(* IEC 61131-3 sources: daoli-st-library/DL_Device (part 25) *)

(* ---- FB_DL_IvBcdExport.st ---- *)
(*==============================================================================
 * 组件名称 (Component)  : FB_DL_IvBcdExport
 * 所属子库 (Sublibrary) : DL_Device
 * 当前版本 (Version)    : 1.0.0
 * 兼容性   (Platform)   : CODESYS 3.5+ / TwinCAT 3 / 汇川 InoProShop / 施耐德 Machine Expert
 *                         仅依赖 Standard.library（TON / R_TRIG），零厂商私有库
 * 功能描述 (Function)   : IV 测试仪 BCD 拨码设定导出。
 *                         把上位下发的十进制设定值（0..9999）拆成四位十进制数字，打包成 BCD 字，
 *                         经"导出脉冲 → 等回读 → 逐位比对"的握手闭环确认测试仪已正确接收；
 *                         回读不一致或超时即锁存故障，等人工复位后重导。
 *                         **面板互转语义（双向，写死）**：
 *                           正解：value → 四位数字 d1(个)…d4(千) → uBcd = d4·16#1000 + d3·16#0100 + d2·16#0010 + d1
 *                           反解：uBcd → value（用于回读通道是 BCD 字的机型，本件按整值比对不拆位）
 *                         两位以上的半字节合法性由"十进制拆分"结构性保证（每位恒 0..9），
 *                         故不存在"非 BCD 半字节"可导出；真正的越界风险在**设定值本身越域**，
 *                         故设 0..9999 域闸 + 越域拒导出（eRangeBad，信息级，不锁存）。
 *                         验收向量：
 *                           ① 设定 1234 → 数字 d1=4, d2=3, d3=2, d4=1；uBcd = 16#1234
 *                           ② 设定 0    → 数字全 0；uBcd = 16#0000（合法边界，不拒算）
 *                           ③ 设定 9999 → uBcd = 16#9999（上界，不溢出）
 *                           ④ 设定 10000 → 拒导出 + eRangeBad（域闸，信息级）
 *                           ⑤ 回读 = 16#1234 → bReadbackOk；回读 = 16#1235 → 锁存 eRbMismatch
 * 接口     (Interface)  : 入 iSetValue 设定值、bExport 导出沿、bReadbackValid 回读有效、
 *                         iReadbackBcd 回读 BCD 字、tReadbackTo 回读超时、bReset 复位沿；
 *                         出 uBcdPacked 打包 BCD 字、abDigits 四位数字（1..4 = 个/十/百/千）、
 *                         bExported 导出脉冲（单拍）、bReadbackOk 回读一致脉冲（单拍）、
 *                         bRbFailed 回读失败锁存、eState 相、eCause 成因、bError 故障标志。
 * 边界     (Boundary)   : ① **属主边界（写死）：本件只做"设定值编码 + 导出握手"，不驱动拨码
 *                         继电器/光电隔离板、不解析 IV 测量曲线**（属测试仪通讯件与曲线件）；
 *                         ② **域闸**：iSetValue 越 0..9999 → 拒导出（信息级 eRangeBad，不锁存、
 *                         不改已导出值）；③ **移位量常量化**：打包移位量取常量 0/4/8/12，
 *                         恒小于 WORD 位宽 16，跨平台无未定义行为（R48/R295）；
 *                         ④ **回读超时 TON**：tonRb 段 0 无条件调用，IN 串 (NOT _bFault)，
 *                         故障期不累计，复位同拍不会立即重锁（R252）；
 *                         ⑤ **锁存解除式**：bRbFailed 与 eFault 仅由 bReset 上升沿解除
 *                         （R228B 唯一迁出），bReset 为外部引脚、恒可达；
 *                         ⑥ **握手单拍脉冲三律**：导出脉冲与回读成功脉冲均在 CASE 内用内部位
 *                         置位、段尾统一映射出口，禁同相内置位后同相撤位（R129）；
 *                         ⑦ 零全局耦合、零物理地址。
 * 分工声明 (Scope)      : 本件只管"设定值 BCD 导出与回读校验"。不接管：花篮标签打印联动
 *                         （属 FB_DL_CassetteBcdLabel）、纯数值 BCD 转换原子件（属 FC_DL_WordToBcd 族）、
 *                         IV 量测流程（属测试顺控件）。
 * 来源标签 (Source Tag) : ROADMAP 空勾真缺口 P2（BCD 设定导出，自研 clean-room）
 * 码表     (Codes)      : 本件不占用任何全局数字码位（零码位范式 R297）；诊断由 BOOL + ENUM 出口承担。
 * 红线自检 (Redline)    : R1 ✓ 零 GVL/VAR_EXTERNAL ｜ R2 ✓ 零 %I/%Q/%M ｜ R3 ✓ 纯 IEC 61131-3
 *                         R4 ✓ 域闸 + 常量移位 + 超时 TON + 单拍脉冲两段式 ｜ R5 ✓ 声明逐行同行双语注释
 *                         R6 ✓ ENUM+CASE 含 ELSE 兜底 ｜ R7 ✓ TON/R_TRIG 段 0 无条件刷新
 * 修订历史 (Revision)   : 2026-11-19  v1.0.0  R47 首版（批次 2 · 序号 10）
 *==============================================================================*)

TYPE E_DL_IbeState :
(
    eIdle    := 0,    // 待机相（可接受导出请求） / Idle, ready for an export request
    eWaitRead:= 10,   // 等回读相（握手窗口内） / Waiting for the read-back
    eFault   := 90    // 故障相（等复位） / Fault, awaiting reset
);
END_TYPE

TYPE E_DL_IbeCause :
(
    eNone       := 0,   // 无异常 / No anomaly
    eRangeBad   := 1,   // 设定值越 0..9999（信息级，拒导出） / Set point out of 0..9999, info level
    eRbMismatch := 2,   // 回读不一致（锁存，故障级） / Read-back mismatch, latched, fault level
    eRbTimeout  := 3,   // 回读超时（锁存，故障级） / Read-back timeout, latched, fault level
    eCfgIllegal := 4,   // 组态非法（超时非正） / Illegal configuration, non-positive timeout
    ePhaseBad   := 5    // 非法相位兜底 / Illegal phase fallback
);
END_TYPE

FUNCTION_BLOCK FB_DL_IvBcdExport
VAR_INPUT
    iSetValue     : INT := 0;              // 设定值，域 0..9999 [-] / Set point, domain 0..9999
    bExport       : BOOL := FALSE;         // 导出请求沿 [-] / Export request edge
    bReadbackValid: BOOL := FALSE;         // 回读有效（当拍电平） [-] / Read-back valid, level
    iReadbackBcd  : INT := 0;              // 回读 BCD 字（按整值比对） [BCD] / Read-back BCD word, compared as a whole
    tReadbackTo   : TIME := T#2S;          // 回读超时，域 > T#0S [ms] / Read-back timeout, > T#0S
    bReset        : BOOL := FALSE;         // 故障复位沿 [-] / Fault reset edge
END_VAR
VAR_OUTPUT
    uBcdPacked  : WORD := 16#0000;                       // 打包 BCD 字（千/百/十/个） [BCD] / Packed BCD word
    abDigits    : ARRAY[1..4] OF BYTE;                   // 四位十进制数字（1=个,2=十,3=百,4=千） [-] / Four decimal digits
    bExported   : BOOL := FALSE;                         // 导出脉冲（单拍） [-] / Export pulse, single scan
    bReadbackOk : BOOL := FALSE;                         // 回读一致脉冲（单拍） [-] / Read-back match pulse, single scan
    bRbFailed   : BOOL := FALSE;                         // 回读失败锁存（等复位） [-] / Read-back failure, latched
    eState      : E_DL_IbeState := E_DL_IbeState.eIdle;  // 相出口 [-] / Phase outlet
    eCause      : E_DL_IbeCause := E_DL_IbeCause.eNone;  // 成因出口（R190 归因唯一） [-] / Cause outlet
    bError      : BOOL := FALSE;                         // 故障标志（仅故障级成因） [-] / Error flag, fault level only
END_VAR
VAR
    _eState   : E_DL_IbeState := E_DL_IbeState.eIdle;    // 内部相（CASE 唯一写入目标） / Internal phase
    _eCause   : E_DL_IbeCause := E_DL_IbeCause.eNone;    // 成因锁存量 / Latched cause
    _bFault   : BOOL := FALSE;                           // 故障锁存位 / Latched fault bit
    _bRbFail  : BOOL := FALSE;                           // 回读失败锁存位 / Latched read-back failure
    _iWork    : INT := 0;                                // 十进制拆分工作值 [-] / Decimal split working value
    _uBcd     : WORD := 16#0000;                         // 打包工作值 [BCD] / Packing working value
    _iRbExp   : INT := 0;                                // 期望回读值（导出时的 BCD 整值） [BCD] / Expected read-back value
    _bExported: BOOL := FALSE;                           // 导出脉冲内部位（单拍） / Internal export pulse
    _bRbOk    : BOOL := FALSE;                           // 回读成功内部位（单拍） / Internal read-back OK pulse
    _bCfgBad  : BOOL := FALSE;                           // 组态非法当拍量 / Illegal configuration this scan
    tonRb     : TON;                                     // 回读超时实例，段 0 无条件调用 / Read-back timeout instance
    rtExport  : R_TRIG;                                  // 导出沿实例，段 0 无条件调用 / Export edge instance
    rtReset   : R_TRIG;                                  // 复位沿实例，段 0 无条件调用 / Reset edge instance
END_VAR
VAR CONSTANT
    DL_IBE_MAX  : INT := 9999;            // 设定值上限（四位十进制） [-] / Set-point upper bound
    DL_IBE_SH0  : WORD := 16#0000;        // 个位打包基准（占位常量，便于口径统一） [BCD] / Units packing base
    DL_IBE_SH4  : INT := 4;               // 十位左移量（恒 < 16，R48） [bit] / Tens shift, always below 16 bits
    DL_IBE_SH8  : INT := 8;               // 百位左移量（恒 < 16，R48） [bit] / Hundreds shift
    DL_IBE_SH12 : INT := 12;              // 千位左移量（恒 < 16，R48） [bit] / Thousands shift
    DL_IBE_MSK  : WORD := 16#000F;        // 半字节掩码（非事件码，头注释声明） [bit] / Nibble mask, not an event code
END_VAR

(* —— 段 0：组态闸 + TON 与两沿无条件周期刷新（R228A；IN 串故障否决，R252） —— *)
_bCfgBad := (tReadbackTo <= T#0S);                             // 回读超时须为正 / Timeout must be positive
rtExport(CLK := bExport);                                      // 导出沿 / Export edge
rtReset(CLK := bReset);                                        // 复位沿 / Reset edge
tonRb(IN := (_eState = E_DL_IbeState.eWaitRead) AND (NOT _bFault), PT := tReadbackTo);   // 回读超时（等回读相派生） / Read-back timeout

(* —— 段 1：单拍量预清零（锁存量 _eCause/_bFault/_bRbFail/_iRbExp 不入清单，R107） —— *)
_bExported := FALSE;                                           // 导出脉冲预清 / Export pulse preset
_bRbOk     := FALSE;                                           // 回读成功脉冲预清 / Read-back OK pulse preset
bError     := FALSE;                                           // 故障标志预清（R45 配对） / Error preset

(* —— 段 2：组态闸（非法即锁存故障级） —— *)
IF _bCfgBad THEN
    _eCause := E_DL_IbeCause.eCfgIllegal;                       // 归因：组态非法 / Cause: illegal configuration
    _bFault := TRUE;                                            // 锁存 / Latch
    _eState := E_DL_IbeState.eFault;                            // 入故障相 / Enter fault phase
END_IF

(* —— 段 3：迁出链（bReset 上升沿：清故障与回读失败锁存，R228B） —— *)
IF rtReset.Q THEN
    _bFault  := FALSE;                                          // 清故障锁存 / Clear fault latch
    _bRbFail := FALSE;                                          // 清回读失败锁存 / Clear read-back failure latch
    _eCause  := E_DL_IbeCause.eNone;                            // 清成因 / Clear cause
    _eState  := E_DL_IbeState.eIdle;                            // 回待机相 / Back to idle
END_IF

(* —— 段 4：相迁移（导出 / 回读握手闭环） —— *)
IF (NOT _bFault) AND (NOT _bCfgBad) THEN
    CASE _eState OF

    E_DL_IbeState.eIdle:
        IF rtExport.Q THEN
            IF (iSetValue < 0) OR (iSetValue > DL_IBE_MAX) THEN
                _eCause := E_DL_IbeCause.eRangeBad;              // 域闸：越域拒导出（信息级，不锁存） / Out of range, info level
            ELSE
                (* 十进制拆分（每位恒 0..9，半字节合法由构造保证） *)
                _iWork := iSetValue;                             // 取设定值 / Take the set point
                abDigits[1] := INT_TO_BYTE(_iWork MOD 10);       // 个位 / Units
                _iWork := _iWork / 10;                           // 去掉个位 / Drop the units digit
                abDigits[2] := INT_TO_BYTE(_iWork MOD 10);       // 十位 / Tens
                _iWork := _iWork / 10;                           // 去掉十位 / Drop the tens digit
                abDigits[3] := INT_TO_BYTE(_iWork MOD 10);       // 百位 / Hundreds
                _iWork := _iWork / 10;                           // 去掉百位 / Drop the hundreds digit
                abDigits[4] := INT_TO_BYTE(_iWork MOD 10);       // 千位 / Thousands

                (* 打包 BCD：移位量为常量，跨平台安全（R48/R295） *)
                _uBcd := SHL(BYTE_TO_WORD(abDigits[4]), DL_IBE_SH12)
                      OR SHL(BYTE_TO_WORD(abDigits[3]), DL_IBE_SH8)
                      OR SHL(BYTE_TO_WORD(abDigits[2]), DL_IBE_SH4)
                      OR (BYTE_TO_WORD(abDigits[1]) AND DL_IBE_MSK);
                uBcdPacked := _uBcd;                             // 打包字出口 / Packed word outlet
                _iRbExp := WORD_TO_INT(_uBcd);                   // 期望回读值（整值比对） / Expected read-back
                _bExported := TRUE;                              // 导出脉冲（内部位，段 7 映射） / Internal export pulse
                _eState := E_DL_IbeState.eWaitRead;              // 进等回读相 / Enter the wait-read phase
            END_IF
        END_IF

    E_DL_IbeState.eWaitRead:
        IF bReadbackValid THEN
            IF iReadbackBcd = _iRbExp THEN
                _bRbOk := TRUE;                                  // 回读一致（内部位） / Read-back matches
                _eState := E_DL_IbeState.eIdle;                  // 回待机相 / Back to idle
            ELSE
                _bRbFail := TRUE;                                // 回读不一致：锁存 / Mismatch: latch
                _bFault  := TRUE;                                // 故障锁存 / Latch the fault
                _eCause  := E_DL_IbeCause.eRbMismatch;           // 归因：回读不一致 / Cause: read-back mismatch
                _eState  := E_DL_IbeState.eFault;                // 入故障相 / Enter fault phase
            END_IF
        ELSIF tonRb.Q THEN
            _bRbFail := TRUE;                                    // 回读超时：锁存 / Timeout: latch
            _bFault  := TRUE;                                    // 故障锁存 / Latch the fault
            _eCause  := E_DL_IbeCause.eRbTimeout;                // 归因：回读超时 / Cause: read-back timeout
            _eState  := E_DL_IbeState.eFault;                    // 入故障相 / Enter fault phase
        END_IF

    E_DL_IbeState.eFault:
        ;                                                        // 故障相：仅等复位沿 / Wait for the reset edge only

    ELSE
        _eCause := E_DL_IbeCause.ePhaseBad;                      // 归因：非法相位 / Cause: illegal phase
        _bFault := TRUE;                                         // 锁存 / Latch
        _eState := E_DL_IbeState.eFault;                         // 强拉故障相 / Force fault phase

    END_CASE
END_IF

(* —— 段 5：出口单点映射（名实双出口，R191） —— *)
bExported   := _bExported;                                       // 导出脉冲出口 / Export pulse outlet
bReadbackOk := _bRbOk;                                           // 回读成功脉冲出口 / Read-back OK outlet
bRbFailed   := _bRbFail;                                         // 回读失败出口 / Read-back failure outlet
eState      := _eState;                                          // 相出口 / Phase outlet
eCause      := _eCause;                                          // 成因出口 / Cause outlet
bError      := _bFault;                                          // 故障标志 / Error flag

END_FUNCTION_BLOCK

(* ---- FB_DL_JunctionBoxPottingCheck.st ---- *)
(*
  FB_DL_JunctionBoxPottingCheck  —  接线盒灌胶量与固化判定 / Junction box potting quantity and cure check
  分类 Category : DL_Device
  码位 Code     : 16#03_2_14
  段位说明      : 03_2 段低半字节 00~0F 已满（05 为历史空穴留存），进位 14 段续号（R192）
  版本 Version  : 1.0.0
  来源 Source   : t2-1-lgf-technology — IEC 61131-3 标准语义的道莅防御性实现
  溯源 Origin   : clean-room 实现，灌胶积分与固化当量公开工艺语义，未复制任何源码行
                  （积分用内部等价实现承载 FB_DL_Integrator 语义；温度域契约对齐 I_DL_TemperatureZone）
  功能 Function : 1) 灌胶量 = 流量对时间积分（DL_TICK 节拍窗离散积分）得 mL，与 fGlueTargetMl ± fGlueTolPct 比较；
                  2) 固化当量 = Σ(max(T − fCureTempMinC, 0) × Δt) 累积 [°C·min]，达 fCureDoseMinCmin 判固化完成；
                  3) 灌胶判据与固化判据独立记账：bGlueOk / bCureOk 不互相覆盖，bCycleOk 仅在两者皆真时为真。
  边界 Boundary : ① fGlueFlowLpm < 0（负流量 = 倒吸）判传感器故障置码进 Fault；
                  ② fGlueTargetMl <= 0 / fCureDoseMinCmin <= 0 / fCureTempMaxC <= fCureTempMinC / 容差 <= 0 判组态错
                     （fCureTempMinC 高于环境上限将永不固化，规格强制）；
                  ③ 超 tCureMax 置 bCureOk := FALSE 并进 Fault（固化超时升级）；
                  ④ 积分节拍窗 DL_TICK 内恒定流量近似（离散积分语义，头注释声明）；
                  ⑤ 解除式自证：Fault 解除 = bReset AND bCycleStart 新上升沿（eState 回 Dose，引脚可满足）；
                  ⑥ CASE 全态覆盖 + ELSE 兜底置故障相。
  依赖 Depends  : I_DL_TemperatureZone（注入，只读属性，不实例化）；积分语义对齐 FB_DL_Integrator（已注册，不实例化）
  码表 Error codes（本件格 03_2_14，子码步进 +0x100）:
    16#0003_0114 信息级：灌胶量达标，Dose 相切换至 Cure 相
    16#0003_0214 故障级：组态非法（目标量/当量下限 <= 0 / 温域倒置 / 容差 <= 0），锁存至复位
    16#0003_0314 故障级：负流量（倒吸）传感器故障，锁存至复位
    16#0003_0414 故障级：固化超时 tCureMax（bCureOk = FALSE）
    16#0003_0514 故障级：状态机落 ELSE 兜底（非法相位 ID）

  修订历史 Revision :
    2026-11-18  v1.0.0  R38 首版
*)

TYPE E_DL_PottingState :
(
    eDose  := 0,    // 灌胶相：流量积分进行中 / Dose, flow integrating
    eCure  := 10,   // 固化相：当量累积进行中 / Cure, equivalent accumulating
    eDone  := 20,   // 完成相：双判据落定 / Done, both verdicts settled
    eFault := 90    // 故障相：组态/倒吸/超时锁定 / Fault, latched
);
END_TYPE

FUNCTION_BLOCK FB_DL_JunctionBoxPottingCheck
VAR_INPUT
    bCycleStart    : BOOL := FALSE;       // 周期启动（上升沿）/ Cycle start
    fGlueFlowLpm   : REAL := 0.0;         // 灌胶流量 [L/min] / Glue flow rate
    fGlueTargetMl  : REAL := 50.0;        // 灌胶目标量 [mL]，域 > 0 / Target dosed volume
    fGlueTolPct    : REAL := 5.0;         // 灌胶容差 [%]，域 > 0 / Dose tolerance
    fCureTempMinC  : REAL := 25.0;        // 固化有效温度下限 [°C] / Cure effective temperature floor
    fCureTempMaxC  : REAL := 80.0;        // 环境/工艺温度上限 [°C]，须 > 下限 / Ambient ceiling, must exceed floor
    fCureDoseMinCmin : REAL := 500.0;     // 固化当量下限 [°C·min]，域 > 0 / Cure equivalent floor
    tCureMax       : TIME := T#3600S;     // 固化最长时限 [ms]，域 > 0 / Cure maximum duration
    bReset         : BOOL := FALSE;       // 复位（Fault 解除路径之一）/ Reset
END_VAR
VAR_OUTPUT
    fGlueDosedMl   : REAL;                // 灌胶量 [mL] / Dosed volume
    fCureDoseCmin  : REAL;                // 固化当量 [°C·min] / Cure equivalent
    bGlueOk        : BOOL;                // 灌胶判据（独立记账）/ Glue verdict, independent bookkeeping
    bCureOk        : BOOL;                // 固化判据（独立记账）/ Cure verdict, independent bookkeeping
    bCycleOk       : BOOL;                // 周期合格（两者皆真）/ Cycle ok, both true
    nErrId         : UDINT;               // 事件码，0 = 无事件 / Event code
    eState         : E_DL_PottingState;   // 状态出口，段尾单点映射 / State outlet
END_VAR
VAR_IN_OUT
    iTempZone : I_DL_TemperatureZone;     // 温区引用（注入，只读属性）/ Temperature zone reference
END_VAR
VAR
    tonTick    : TON;                     // 积分节拍窗，自复位（段 0 无条件刷新）/ Integration tick window, self-resetting
    tonCure    : TON;                     // 固化超时计时，段 0 无条件刷新 / Cure timeout timer
    tonFaultWch: TON;                     // 故障观察窗，自复位 / Fault watch window, self-resetting
    rtStart    : R_TRIG;                  // 周期启动上升沿 / Cycle start rising edge
    rtReset    : R_TRIG;                  // 复位上升沿 / Reset rising edge
    _bTickBrk  : BOOL;                    // 节拍窗断输入请求（自复位范式，R182 同族）/ Tick break request
    _eState    : E_DL_PottingState := E_DL_PottingState.eDose;   // 内部相位（CASE 唯一写入目标）/ Internal phase
    _rTempC    : REAL;                    // 温区实测温度 [°C] / Zone actual temperature
    _rVolRate  : REAL;                    // 流量换算暂存 [mL/s] / Volume rate scratch
    _rTolMl    : REAL;                    // 容差换算暂存 [mL] / Tolerance scratch
    _uFault    : UDINT;                   // 故障码锁存 / Latched fault code
    _uInfo     : UDINT;                   // 信息码，每拍重算 / Info code
    _bFault    : BOOL;                    // 故障锁存位 / Latched fault bit
    _bCfgBad   : BOOL;                    // 组态非法聚合 / Configuration invalid aggregate
    _bGlueHold : BOOL;                    // 灌胶判据保持量（独立记账）/ Glue verdict held quantity
    _bCureHold : BOOL;                    // 固化判据保持量（独立记账）/ Cure verdict held quantity
    _bCureMax  : BOOL;                    // 固化超时保持量 / Cure timeout held quantity
END_VAR
VAR CONSTANT
    DL_TICK    : TIME := T#100MS;   // 积分节拍窗 [ms]（离散积分步长）/ Integration tick window
    DL_LPM2MLS : REAL := 16.6667;   // L/min → mL/s 换算系数 / Litres-per-minute to mL-per-second factor
    rFinLim    : REAL := 1.0E15;    // 非有限值筛查幅值上限 / Non-finite screening cap
    DL_WatchPt : TIME := T#2S;      // 故障观察窗 [ms]，自复位 / Fault watch window
END_VAR

(* —— 段 0：定时器与边沿无条件周期刷新（R182：调用语句不得置于 IF/CASE 内） —— *)
rtStart(CLK := bCycleStart);                                    // 周期启动上升沿，每拍必调
rtReset(CLK := bReset);                                         // 复位上升沿，每拍必调
tonFaultWch(IN := (NOT tonFaultWch.Q), PT := DL_WatchPt);       // 观察窗自复位（表达式入参）
tonTick(IN := (NOT tonTick.Q) AND (NOT _bTickBrk), PT := DL_TICK);   // 节拍窗自复位（表达式入参，禁外部沿清零）
_bTickBrk := FALSE;                                             // 断输入拍在调用后自清（R188 范式）
tonCure(IN := (_eState = E_DL_PottingState.eCure), PT := tCureMax);  // 固化超时（表达式入参，相位条件不写进 IF）

(* —— 段 1：单拍量预清零（锁存量 _uFault/_bFault/_bGlueHold/_bCureHold/_bCureMax/_rVolRate 不入清单，R187①） —— *)
_uInfo := 16#0000_0000;         // 信息码每拍重算
_bCfgBad := FALSE;              // 组态非法预清零
nErrId := 16#0000_0000;         // 事件码缺省无事件

(* —— 段 2：组态域闸（覆盖全部参与判据换算的引脚，R151） —— *)
IF (fGlueTargetMl <> fGlueTargetMl) OR (fGlueTargetMl <= 0.0) OR (ABS(fGlueTargetMl) > rFinLim) THEN
    _bCfgBad := TRUE;           // 目标量非法
END_IF
IF (fGlueTolPct <= 0.0) OR (fCureDoseMinCmin <= 0.0) THEN
    _bCfgBad := TRUE;           // 容差/当量下限非法（防除零）
END_IF
IF fCureTempMaxC <= fCureTempMinC THEN
    _bCfgBad := TRUE;           // 温域倒置：固化下限高于环境上限将永不固化（规格强制）
END_IF
IF TIME_TO_DINT(tCureMax) <= 0 THEN
    _bCfgBad := TRUE;           // 超时非法
END_IF

(* —— 段 3：复位沿（Fault 解除式：bReset，eState 回 Dose 等新上升沿） —— *)
IF rtReset.Q THEN
    IF (NOT _bCfgBad) THEN
        _bFault := FALSE;       // 清故障锁存位
        _uFault := 16#0000_0000;
        _eState := E_DL_PottingState.eDose;   // 回灌胶相（等 bCycleStart 新上升沿）
    END_IF
END_IF

(* —— 段 4：温区只读采集 + 节拍窗离散积分（窗内恒定近似，头注释声明） —— *)
_rTempC := iTempZone.fTempActual;       // 实测温度 [°C]（只读属性）
IF tonTick.Q THEN
    _bTickBrk := TRUE;                  // 断输入请求：下一拍窗重开（自复位范式）
    _rVolRate := fGlueFlowLpm * DL_LPM2MLS;                  // [mL/s]（负值即倒吸，段 5 判）
    fGlueDosedMl := fGlueDosedMl + _rVolRate * (TIME_TO_REAL(DL_TICK) / 1000.0);   // 流量积分 [mL]
    fCureDoseCmin := fCureDoseCmin + MAX(_rTempC - fCureTempMinC, 0.0)
                     * (TIME_TO_REAL(DL_TICK) / 60000.0);                     // 当量积分 [°C·min]
END_IF

(* —— 段 5：相位机（只做迁移与判据记账；出口在段 8） —— *)
CASE _eState OF

E_DL_PottingState.eDose:
    IF _bCfgBad THEN
        _uFault := 16#0003_0214;        // 故障级：组态非法
        _bFault := TRUE;                // 锁存（复位沿可清）
        _eState := E_DL_PottingState.eFault;
    ELSIF fGlueFlowLpm < 0.0 THEN
        _uFault := 16#0003_0314;        // 故障级：负流量倒吸（传感器故障）
        _bFault := TRUE;
        _eState := E_DL_PottingState.eFault;
    ELSE
        _rTolMl := fGlueTargetMl * fGlueTolPct / 100.0;     // 容差 [mL]
        IF fGlueDosedMl >= (fGlueTargetMl - _rTolMl) THEN
            IF fGlueDosedMl <= (fGlueTargetMl + _rTolMl) THEN
                _bGlueHold := TRUE;     // 灌胶判据记账：达标（独立，不覆盖固化）
                _uInfo := 16#0003_0114; // 信息级：灌胶量达标
            ELSE
                _bGlueHold := FALSE;    // 过量超容差：判不合格
            END_IF
            _eState := E_DL_PottingState.eCure;   // 切固化相（量已定，不再积分判定）
        END_IF
    END_IF

E_DL_PottingState.eCure:
    IF fCureDoseCmin >= fCureDoseMinCmin THEN
        _bCureHold := TRUE;             // 固化判据记账：达标（独立，不覆盖灌胶）
        _eState := E_DL_PottingState.eDone;   // 进完成相
    ELSIF tonCure.Q THEN
        _uFault := 16#0003_0414;        // 故障级：固化超时（bCureOk = FALSE，规格强制）
        _bFault := TRUE;
        _bCureHold := FALSE;            // 固化判据显式记账为不合格
        _eState := E_DL_PottingState.eFault;
    END_IF

E_DL_PottingState.eDone:
    ;                                   // 完成相：判据已落定，等新周期（bCycleOk 段 8 出口）

E_DL_PottingState.eFault:
    ;                                   // 故障相：等复位沿（段 3 承载解除）

ELSE
    _uFault := 16#0003_0514;            // 故障级：非法相位 ID 兜底
    _bFault := TRUE;                    // 锁存
    _eState := E_DL_PottingState.eFault;// 强制回故障相

END_CASE

(* —— 段 7：出口单点映射（名实同源；独立记账，禁互相覆盖） —— *)
bGlueOk  := _bGlueHold AND (NOT _bCfgBad);      // 灌胶判据出口（独立）
bCureOk  := _bCureHold AND (NOT _bCfgBad);      // 固化判据出口（独立）
bCycleOk := bGlueOk AND bCureOk;                // 周期合格：两者皆真
IF _bCfgBad THEN
    nErrId := 16#0003_0214;         // 故障级：组态非法（每拍重申，复位沿清）
    _bFault := TRUE;
ELSIF fGlueFlowLpm < 0.0 THEN
    nErrId := 16#0003_0314;         // 故障级：负流量（锁存语义由 Fault 相承载）
    _bFault := TRUE;
END_IF
IF _bFault THEN
    nErrId := _uFault;              // 故障锁存码回放（不在故障相按当下输入重推）
    bGlueOk  := FALSE;              // 故障相判据出口撤销（安全侧）
    bCureOk  := FALSE;
    bCycleOk := FALSE;
END_IF
eState := _eState;                  // 状态出口单点映射

END_FUNCTION_BLOCK

(* ---- FB_DL_KilnPreheatStageSeq.st ---- *)
(*
  DL Factory R84 | FB_DL_KilnPreheatStageSeq
  功能：预热器旋风级联投料时序，含各级压差确认、堵料判据与喂料升速
  开源溯源：无（clean-room 自研，依据公开工艺公式，来源=行业通用公式，许可证=MIT，借鉴点=公式结构）
  规则：R1-R16 全遵守
*)
TYPE E_DL_KilnPreState :
(
    eIdle := 0, // 空闲待启动 [-] / idle [-]
    eStageCheck := 1, // 各级压差确认相 [-] / stage pressure check phase [-]
    eFeedOn := 2, // 喂料投入相 [-] / feed on phase [-]
    eStableCheck := 3, // 稳定确认相 [-] / stability confirmation phase [-]
    eFeedUp := 4, // 喂料升速相 [-] / feed ramp up phase [-]
    eDone := 5, // 完成相 [-] / done phase [-]
    eFault := 6 // 故障锁存相 [-] / fault latched phase [-]
) := eIdle;
END_TYPE

FUNCTION_BLOCK FB_DL_KilnPreheatStageSeq
VAR_INPUT
    xStart : BOOL; // 级联投料启动命令 [-] / cascade feed start command [-]
    xReset : BOOL; // 复位命令，上升沿清故障码与堵料位 [-] / reset command [-]
    aStageDpKpa : ARRAY[0..3] OF REAL; // 四级旋风筒压差（C1..C4） [kPa] / stage pressure drops C1 to C4 [kPa]
    fDpMinKpa : REAL := 0.3; // 单级最小压差（低于即判断料不畅） [kPa] / minimum stage pressure drop [kPa]
    fDpBlockKpa : REAL := 2.5; // 单级堵料压差阈值 [kPa] / blockage pressure threshold [kPa]
    xFeedReady : BOOL; // 喂料设备就绪反馈 [-] / feed equipment ready feedback [-]
    fFeedTph : REAL; // 当前喂料量 [t/h] / current feed rate [t/h]
    fFeedTargetTph : REAL := 180.0; // 目标喂料量 [t/h] / target feed rate [t/h]
    fFeedOnTph : REAL := 5.0; // 喂料已投入判据下限 [t/h] / feed on detection floor [t/h]
    tCheckLimit : TIME := T#30S; // 压差确认超时 [s] / pressure check timeout [s]
    tStableLimit : TIME := T#120S; // 稳定确认时长 [s] / stability confirmation duration [s]
    tRampLimit : TIME := T#600S; // 升速相超时 [s] / ramp up timeout [s]
    tScan : TIME := T#100MS; // 扫描周期 [s] / scan period [s]
END_VAR
VAR_OUTPUT
    eState : E_DL_KilnPreState; // 当前时序状态 [-] / current sequence state [-]
    iErrCode : INT; // 故障码 0=正常，701~706 [-] / error code, 701 to 706 [code]
    xBlocked : BOOL; // 堵料标志（锁存至复位沿） [-] / blockage flag latched [-]
    xDone : BOOL; // 完成单拍脉冲 [-] / done one-shot pulse [-]
END_VAR
VAR
    rtStart : R_TRIG; // 启动上升沿实例 [-] / start rising edge instance [-]
    rtReset : R_TRIG; // 复位上升沿实例 [-] / reset edge instance [-]
    tonCheck : TON; // 压差确认超时定时器 [-] / pressure check timer [-]
    tonFeed : TON; // 喂料投入超时定时器（独立实例，避免与确认相共计时） [-] / feed on timer, a dedicated instance [-]
    tonStable : TON; // 稳定确认定时器 [-] / stability timer [-]
    tonRamp : TON; // 升速相超时定时器 [-] / ramp timeout timer [-]
    _eState : E_DL_KilnPreState := E_DL_KilnPreState.eIdle; // 内部相位（CASE 唯一写目标） [-] / internal phase [-]
    _iErr : INT; // 故障码内部锁存 [-] / latched error code [-]
    _bBlocked : BOOL; // 堵料内部锁存 [-] / internal blockage latch [-]
    xDoneInt : BOOL; // 完成内部锁存位 [-] / internal done latch [-]
    xDonePrev : BOOL; // 完成前拍快照 [-] / done previous scan snapshot [-]
    i : INT; // 级索引游标（0→3 正向） [-] / stage cursor, forward only [-]
    xDpBad : BOOL; // 压差非有限或越界当拍标志 [-] / pressure bad flag [-]
    xBlockNow : BOOL; // 本拍堵料判据 [-] / blockage verdict of this scan [-]
    fStepTph : REAL; // 本拍升速增量 [t/h] / ramp increment of this scan [t/h]
    fDtSec : REAL; // 扫描周期秒值 [s] / scan period in seconds [s]
END_VAR

// 段 0｜边沿与定时器实例无条件周期刷新（R7）
rtStart(CLK := xStart); // 启动沿每拍必调 [-] / start edge every scan [-]
rtReset(CLK := xReset); // 复位沿每拍必调 [-] / reset edge every scan [-]
tonCheck(IN := _eState = E_DL_KilnPreState.eStageCheck, PT := tCheckLimit); // 确认相独立计时 [-] / check phase timer [-]
tonFeed(IN := _eState = E_DL_KilnPreState.eFeedOn, PT := tCheckLimit); // 喂料相独立计时 [-] / feed on phase timer [-]
tonStable(IN := _eState = E_DL_KilnPreState.eStableCheck, PT := tStableLimit); // 稳定相闸 [-] / stability gate [-]
tonRamp(IN := _eState = E_DL_KilnPreState.eFeedUp, PT := tRampLimit); // 升速相闸 [-] / ramp gate [-]

// 段 1｜四级压差异常与堵料判据（定长数组，正向游标 0→3）
fDtSec := LREAL_TO_REAL(TIME_TO_LREAL(tScan) / 1000.0); // ms ÷ 1000 = s / [ms] / 1000 = [s]
xDpBad := FALSE; // 初值置假 [-] / start false [-]
xBlockNow := FALSE; // 初值置假 [-] / start false [-]
FOR i := 0 TO 3 DO
    IF NOT (aStageDpKpa[i] > -1.0E30 AND aStageDpKpa[i] < 1.0E30) THEN
        xDpBad := TRUE; // 压差非有限（变送器失效） [-] / non finite pressure drop [-]
    ELSIF aStageDpKpa[i] > fDpBlockKpa THEN
        xBlockNow := TRUE; // 单级压差超堵料阈值 [-] / stage pressure above the blockage threshold [-]
    END_IF
END_FOR
IF xBlockNow THEN
    _bBlocked := TRUE; // 堵料锁存（复位沿清） [-] / latch the blockage, cleared on reset [-]
END_IF

// 段 2｜复位沿：清故障码、堵料位与相位（R189）
IF rtReset.Q THEN
    _iErr := 0; // 清故障码 [-] / clear error code [-]
    _bBlocked := FALSE; // 清堵料锁存 [-] / clear the blockage latch [-]
    xDoneInt := FALSE; // 清完成锁存 [-] / clear done latch [-]
    _eState := E_DL_KilnPreState.eIdle; // 回空闲相 [-] / back to idle [-]
END_IF

// 段 3｜主状态机（合法事件优先于超时迁移，R275）
CASE _eState OF
    E_DL_KilnPreState.eIdle: // 空闲相 [-] / idle [-]
        xDoneInt := FALSE; // 空闲清完成锁存 [-] / clear done latch in idle [-]
        IF rtStart.Q THEN
            _eState := E_DL_KilnPreState.eStageCheck; // 启动沿进压差确认相 [-] / start edge enters the check [-]
        END_IF
    E_DL_KilnPreState.eStageCheck: // 各级压差确认相 [-] / stage pressure check [-]
        IF xBlockNow THEN
            _iErr := 701; _eState := E_DL_KilnPreState.eFault; // 投料前已堵料 [-] / blockage before feeding [-]
        ELSIF xDpBad THEN
            _iErr := 702; _eState := E_DL_KilnPreState.eFault; // 压差信号失效 [-] / pressure signal invalid [-]
        ELSIF tonCheck.Q THEN
            _iErr := 703; _eState := E_DL_KilnPreState.eFault; // 压差建立超时（通风不足） [-] / pressure build up timeout [-]
        ELSIF (aStageDpKpa[0] >= fDpMinKpa) AND (aStageDpKpa[1] >= fDpMinKpa) AND (aStageDpKpa[2] >= fDpMinKpa) AND (aStageDpKpa[3] >= fDpMinKpa) THEN
            _eState := E_DL_KilnPreState.eFeedOn; // 各级压差均达标转喂料相 [-] / all stages above the floor leads to feed on [-]
        END_IF
    E_DL_KilnPreState.eFeedOn: // 喂料投入相 [-] / feed on [-]
        IF NOT xFeedReady THEN
            _iErr := 704; _eState := E_DL_KilnPreState.eFault; // 喂料设备未就绪 [-] / feed equipment not ready [-]
        ELSIF xDpBad THEN
            _iErr := 702; _eState := E_DL_KilnPreState.eFault; // 喂料中压差信号失效（R583 补：原仅两相有闸） [-] / pressure signal lost while feeding [-]
        ELSIF xBlockNow THEN
            _iErr := 701; _eState := E_DL_KilnPreState.eFault; // 投料中堵料 [-] / blockage while feeding [-]
        ELSIF fFeedTph >= fFeedOnTph THEN
            _eState := E_DL_KilnPreState.eStableCheck; // 喂料已建立转稳定确认 [-] / feed established leads to stability check [-]
        ELSIF tonFeed.Q THEN
            _iErr := 705; _eState := E_DL_KilnPreState.eFault; // 喂料未建立超时 [-] / feed on timeout [-]
        END_IF
    E_DL_KilnPreState.eStableCheck: // 稳定确认相 [-] / stability check [-]
        IF xBlockNow THEN
            _iErr := 701; _eState := E_DL_KilnPreState.eFault; // 稳定期堵料 [-] / blockage during the stability window [-]
        ELSIF xDpBad THEN
            _iErr := 702; _eState := E_DL_KilnPreState.eFault; // 压差信号失效 [-] / pressure signal invalid [-]
        ELSIF tonStable.Q THEN
            _eState := E_DL_KilnPreState.eFeedUp; // 稳定时长满转升速相 [-] / stable window elapsed leads to ramp up [-]
        END_IF
    E_DL_KilnPreState.eFeedUp: // 喂料升速相 [-] / feed ramp up [-]
        fStepTph := 0.5 * fDtSec; // (t/h)/s × s = t/h（固定 0.5 t/h 每秒升幅） / [t/h] per [s] × [s] = [t/h]
        IF xDpBad THEN
            _iErr := 702; _eState := E_DL_KilnPreState.eFault; // 升速中压差信号失效（R583 补） [-] / pressure signal lost during ramp up [-]
        ELSIF xBlockNow THEN
            _iErr := 701; _eState := E_DL_KilnPreState.eFault; // 升速中堵料（立即停止喂料） [-] / blockage during ramp up [-]
        ELSIF (fFeedTargetTph - fFeedTph) <= fStepTph THEN
            _eState := E_DL_KilnPreState.eDone; // 达目标喂料量转完成相 [-] / target reached leads to done [-]
        ELSIF tonRamp.Q THEN
            _iErr := 705; _eState := E_DL_KilnPreState.eFault; // 升速超时（未达目标） [-] / ramp up timeout [-]
        END_IF
    E_DL_KilnPreState.eDone: // 完成相 [-] / done [-]
        xDoneInt := TRUE; // 置完成锁存（出口统一映射单拍） [-] / raise done latch [-]
        IF NOT xStart THEN
            _eState := E_DL_KilnPreState.eIdle; // 命令撤销回空闲 [-] / command released returns to idle [-]
        END_IF
    E_DL_KilnPreState.eFault: // 故障相：码值锁存回放，仅复位沿出 [-] / fault, exit only on reset [-]
        ; // 锁存回放（R28） [-] / replay the latch only [-]
ELSE
    _iErr := 706; _eState := E_DL_KilnPreState.eFault; // 非法相位兜底 [-] / illegal phase fallback [-]
END_CASE

// 段 4｜出口映射（名实双出口，同源赋值）
eState := _eState; // 状态出口 [-] / state outlet [-]
iErrCode := _iErr; // 故障码出口（锁存值） [-] / error code outlet [-]
xBlocked := _bBlocked; // 堵料位出口（锁存值） [-] / blockage outlet [-]
xDone := xDoneInt AND NOT xDonePrev; // 完成单拍（内部锁存 → 出口映射） [-] / done one-shot [-]
xDonePrev := xDoneInt; // 本拍快照供下拍比较 [-] / snapshot for the next scan [-]
END_FUNCTION_BLOCK

(* ---- FB_DL_LadlePourWeightCtrl.st ---- *)
(*
  Component : FB_DL_LadlePourWeightCtrl
  Category  : DL_Device
  Type      : FB
  Complexity: C2
  VERSION   : v1.0.0
  功能      : 浇包定量浇注控制：ENUM 五态（Idle/Fast/Slow/Done/Fault），快浇到"目标-快浇量"转慢浇，慢浇到"目标-提前量"停浇，称重偏差超差报警。
  开源溯源  : 道莅原创 clean-room 自研（无外部代码引用）｜License: MIT
  边界条件  : ① 目标重量、快浇量、提前量、公差须满足 快浇量 < 目标重量 且公差 > 0，否则拒绝启动并锁故障；
              ② 提前量用于补偿落料惯性，提前量 >= 目标重量时判组态非法（永不达量）；
              ③ 浇注全程有超时监控；偏差百分比在每拍按输入重算（信息量，不入锁存）。
*)

TYPE E_DL_PourPhase :
(
    eIdle  := 0,    (* 空闲：等待启动条件 / Idle waiting start *)
    eFast  := 10,   (* 快浇：大流量阶段 / Fast pouring stage *)
    eSlow  := 20,   (* 慢浇：精计量阶段 / Slow metering stage *)
    eDone  := 50,   (* 完成：偏差已判定 / Done, deviation judged *)
    eFault := 90    (* 故障：锁存待复位 / Fault latched *)
);
END_TYPE

FUNCTION_BLOCK FB_DL_LadlePourWeightCtrl
VAR_INPUT
    bEnable     : BOOL;   (* 使能电平 [-] Enable level *)
    bReset      : BOOL;   (* 复位上升沿，清故障锁存 [-] Reset edge *)
    bStart      : BOOL;   (* 启动上升沿 [-] Start edge *)
    bLadleReady : BOOL;   (* 浇包就位反馈 [-] Ladle in position feedback *)
    fWeightKg   : REAL;   (* 称重实测重量 [kg] Measured weight *)
    fTargetKg   : REAL;   (* 目标浇注重量 [kg] Target pouring weight *)
    fFastToKg   : REAL;   (* 快浇转慢浇的剩余量 [kg] Fast-to-slow switch remainder *)
    fAdvanceKg  : REAL;   (* 停浇提前量（落料惯性补偿） [kg] Stop advance *)
    fTolPct     : REAL;   (* 称重偏差公差 [%] Weight deviation tolerance *)
    tPourTo     : TIME;   (* 浇注全程超时 [ms] Pouring overall timeout *)
END_VAR
VAR_OUTPUT
    bPourFast : BOOL;              (* 快浇阀输出 [-] Fast pour valve output *)
    bPourSlow : BOOL;              (* 慢浇阀输出 [-] Slow pour valve output *)
    fDevPct   : REAL;              (* 相对目标重量偏差 [%] Weight deviation percent *)
    bOverTol  : BOOL;              (* 偏差超差报警 [-] Deviation over tolerance *)
    bDone     : BOOL;              (* 浇注完成（锁存） [-] Pouring done latched *)
    ePhase    : E_DL_PourPhase;    (* 相位出口，段尾单点映射 [-] Phase outlet *)
    bError    : BOOL;              (* 故障锁存标志 [-] Fault latch flag *)
    uErrId    : UDINT;             (* 事件码，0 = 无事件 [-] Event code *)
END_VAR
VAR
    rtReset  : R_TRIG;   (* 复位沿实例，每拍无条件刷新 / Reset edge *)
    rtStart  : R_TRIG;   (* 启动沿实例，每拍无条件刷新 / Start edge *)
    tonPourTo: TON;      (* 浇注全程超时（专用超时件） / Pouring timeout *)
    _ePhase  : E_DL_PourPhase := E_DL_PourPhase.eIdle;  (* 内部相位 / Internal phase *)
    _bFault  : BOOL;     (* 故障锁存位（锁存量） / Latched fault bit *)
    _uFault  : UDINT;    (* 故障码锁存（锁存量） / Latched fault code *)
    _bDone   : BOOL;     (* 完成锁存位（锁存量） / Latched done bit *)
    _bOver   : BOOL;     (* 超差锁存位（锁存量） / Latched over-tolerance bit *)
    _bCfgBad : BOOL;     (* 组态非法当拍量 [-] Config illegal flag *)
    _bNonFin : BOOL;     (* 输入非有限当拍量 [-] Non-finite input flag *)
END_VAR
VAR CONSTANT
    DL_EPS      : REAL := 1.0E-9;   (* 除零判定容差 [无量纲] Divide-by-zero tolerance *)
    DL_PCT_BASE : REAL := 100.0;    (* 百分比基准 [%] Percent base *)
    DL_ZERO     : REAL := 0.0;      (* 零常量 [无量纲] Zero constant *)
END_VAR

(* —— 段 0｜沿与定时器每拍无条件刷新（禁置于 IF/CASE 内，使能挂 IN 引脚） —— *)
rtReset(CLK := bReset);
rtStart(CLK := bStart);
tonPourTo(IN := ((_ePhase = E_DL_PourPhase.eFast) OR (_ePhase = E_DL_PourPhase.eSlow))
              AND (NOT _bFault), PT := tPourTo);

(* —— 段 1｜每拍量预清零（锁存量 _bFault/_uFault/_bDone/_bOver 不入清单） —— *)
uErrId := 16#0000_0000;
_bCfgBad := FALSE;
_bNonFin := FALSE;

(* —— 段 2｜复位沿：一次性清干净（唯一解除路径，恒可达） —— *)
IF rtReset.Q THEN
    _bFault := FALSE;
    _uFault := 16#0000_0000;
    _bDone := FALSE;
    _bOver := FALSE;
    _ePhase := E_DL_PourPhase.eIdle;
END_IF

(* —— 段 3｜非有限拦截与组态闸（覆盖目标/快浇量/提前量/公差/时长） —— *)
IF (fWeightKg <> fWeightKg) OR ((fWeightKg - fWeightKg) <> 0.0)
   OR (fTargetKg <> fTargetKg) OR ((fTargetKg - fTargetKg) <> 0.0)
   OR (fFastToKg <> fFastToKg) OR ((fFastToKg - fFastToKg) <> 0.0)
   OR (fAdvanceKg <> fAdvanceKg) OR ((fAdvanceKg - fAdvanceKg) <> 0.0)
   OR (fTolPct <> fTolPct) OR ((fTolPct - fTolPct) <> 0.0) THEN
    _bNonFin := TRUE;
END_IF
IF (fTargetKg <= DL_EPS) OR (fFastToKg <= DL_ZERO) OR (fFastToKg >= fTargetKg)
   OR (fAdvanceKg < DL_ZERO) OR (fAdvanceKg >= fTargetKg) OR (fTolPct <= DL_ZERO)
   OR (tPourTo = T#0S) THEN
    _bCfgBad := TRUE;
END_IF

(* —— 段 4｜偏差百分比：每拍按输入重算（信息级量，不入锁存） —— *)
IF ABS(fTargetKg) > DL_EPS THEN
    fDevPct := (fWeightKg - fTargetKg) / fTargetKg * DL_PCT_BASE;   (* 分母已过域闸 [%] / Guarded division *)
ELSE
    fDevPct := 0.0;                                (* 目标为 0：偏差无定义，置 0 不留 Inf/NaN / Undefined -> 0 *)
END_IF
IF fDevPct < DL_ZERO THEN
    fDevPct := -fDevPct;                         (* 取绝对值 [%] / Absolute value *)
END_IF

(* —— 段 5｜主状态机：五态全覆盖 + ELSE 兜底 —— *)
CASE _ePhase OF
E_DL_PourPhase.eIdle:
    bPourFast := FALSE; bPourSlow := FALSE;
    IF rtStart.Q AND bEnable AND bLadleReady AND (NOT _bFault)
       AND (NOT _bCfgBad) AND (NOT _bNonFin) THEN
        _bDone := FALSE;
        _bOver := FALSE;
        _ePhase := E_DL_PourPhase.eFast;
    ELSIF rtStart.Q AND (_bFault OR _bCfgBad OR _bNonFin OR (NOT bLadleReady)) THEN
        _bFault := TRUE;                 (* 带病启动拒绝 / Reject start with bad conditions *)
        _uFault := 16#0026_0001;
        _ePhase := E_DL_PourPhase.eFault;
    END_IF

E_DL_PourPhase.eFast:
    bPourFast := TRUE; bPourSlow := FALSE;
    IF _bNonFin THEN
        _bFault := TRUE; _uFault := 16#0026_0002;    (* 故障级：称重非有限 *)
        _ePhase := E_DL_PourPhase.eFault;
    ELSIF fWeightKg >= (fTargetKg - fFastToKg) THEN
        _ePhase := E_DL_PourPhase.eSlow;             (* 迁出条件 1：转慢浇精计量 *)
    ELSIF tonPourTo.Q THEN
        _bFault := TRUE; _uFault := 16#0026_0003;    (* 故障级：快浇超时 *)
        _ePhase := E_DL_PourPhase.eFault;
    ELSIF NOT bEnable THEN
        _ePhase := E_DL_PourPhase.eIdle;             (* 迁出条件 2：使能撤销回安全态 *)
    END_IF

E_DL_PourPhase.eSlow:
    bPourFast := FALSE; bPourSlow := TRUE;
    IF _bNonFin THEN
        _bFault := TRUE; _uFault := 16#0026_0002;    (* 故障级：称重非有限 *)
        _ePhase := E_DL_PourPhase.eFault;
    ELSIF fWeightKg >= (fTargetKg - fAdvanceKg) THEN
        _bDone := TRUE;                              (* 迁出条件 1：到量提前量达成 *)
        _ePhase := E_DL_PourPhase.eDone;
    ELSIF tonPourTo.Q THEN
        _bFault := TRUE; _uFault := 16#0026_0003;    (* 故障级：慢浇超时 *)
        _ePhase := E_DL_PourPhase.eFault;
    ELSIF NOT bEnable THEN
        _ePhase := E_DL_PourPhase.eIdle;             (* 迁出条件 2：使能撤销 *)
    END_IF

E_DL_PourPhase.eDone:
    bPourFast := FALSE; bPourSlow := FALSE;          (* 到量即双阀全关 *)
    IF fDevPct > fTolPct THEN
        _bOver := TRUE;                              (* 超差锁存，待复位清除 *)
    END_IF
    IF NOT bStart THEN
        _ePhase := E_DL_PourPhase.eIdle;             (* 启动撤销：回空闲 *)
    END_IF

E_DL_PourPhase.eFault:
    bPourFast := FALSE; bPourSlow := FALSE;          (* 故障相：双阀全关走安全侧 *)

ELSE
    bPourFast := FALSE; bPourSlow := FALSE;          (* 兜底相：先关双阀再锁故障，安全侧不留上拍开阀值 *)
    _bFault := TRUE;                                 (* 兜底：非法相位锁存 *)
    _uFault := 16#0026_0009;
    _ePhase := E_DL_PourPhase.eFault;
END_CASE

(* —— 段 6｜出口单点映射 —— *)
ePhase := _ePhase;
bDone := _bDone;
bOverTol := _bOver;
bError := _bFault;
IF _bFault AND (_uFault <> 16#0000_0000) THEN
    uErrId := _uFault;                               (* 故障码锁存回放 / Latched fault replay *)
END_IF
END_FUNCTION_BLOCK

(* ---- FB_DL_LamCtrlDualZone.st ---- *)
(*==============================================================================
 * 组件名称 (Component)  : FB_DL_LamCtrlDualZone
 * 所属子库 (Sublibrary) : DL_Device
 * 当前版本 (Version)    : 1.0.0
 * 兼容性 (Platform)     : CODESYS 3.5 / TwinCAT 3 / 汇川 InoProShop（纯标准元素，零方言）
 * 功能描述 (Function)   : 层压机双腔真空协调与差压保护。四段顺控（粗抽→平衡→精抽→
 *                         保压），差压越限时只降抽得快的一侧（双侧同降会把时长翻倍且不
 *                         解决差压）；段超时只报码并保持当前抽速（归零即放弃已有真空度）。
 *                         双腔达标判据为「双侧都不高于目标」。不做泵启停时序、不做阀门
 *                         驱动、不做真空泄漏率诊断（另有专件）。
 * 溯源 (Origin)         : 道莅 clean-room 防御性实现
 * 本文件内含 (Contains) : TYPE E_DL_LamSeg / FUNCTION_BLOCK FB_DL_LamCtrlDualZone
 * 依赖 (Depends)        : 无（仅 Standard.library 的 ABS / MIN / MAX）
 * 红线自检 (Redline)    : 无外部全局变量、无硬件地址直引 ｜ 全变量中英双语同行注释
 *                         差压上限判零防除零 ｜ 目标 ≥ 大气压即组态错 ｜ 单侧非有限按该侧
 *                         0 处理、双侧非有限停车 ｜ 段超时定时器无条件周期刷新 ｜ 枚举显式
 *                         赋值 ｜ CASE 含 ELSE 兜底
 * 错误码表 (Codes)      : 16#0003_03BB 就绪（各段正常或本拍无事件）
 *                         16#0003_03BC 故障级 差压上限 ≤0 或非有限
 *                         16#0003_03BD 故障级 目标真空 ≥ 当地大气压（物理不可达）
 *                         16#0003_03BE 故障级 段超时（保持当前抽速，不归零）
 *                         16#0003_03BF 故障级 单侧真空读数非有限（该侧按 0，双侧齐发即停车）。
 *                                    本件 5 槽全用、无预留槽，已登记待裁定
 * 修订历史 (Revision)   : 2026-11-17  v1.0.0  首版入库 · R28 · 阶段三批 3
 * 验收向量 (Acceptance) : 正向 目标 0.5 kPa、差压上限 3 kPa、上腔 5 / 下腔 12 → 差压 7 越限
 *                         → bDpGuardActive 且降上泵；双腔到 0.5 → bVacOk
 *                         反向 目标设 105 kPa（≥ 大气压）→ 16#0003_03BD；差压上限 0 →
 *                         16#0003_03BC；上腔给 NaN → 16#0003_03BF 且上腔按 0；段拖满 →
 *                         16#0003_03BE 且抽速保持
 *============================================================================*)

(*-----------------------------------------------------------------------------
 * 枚举: E_DL_LamSeg（归属本功能块，同文件发布，全库唯一定义；数值即 uSeg 出口值）
 *----------------------------------------------------------------------------*)
TYPE E_DL_LamSeg :
(
    eIdle    := 0,    // 待机：未启动 / Idle, not started
    eRough   := 1,    // 粗抽：双泵全速 / Rough pumping, both pumps at full speed
    eBalance := 2,    // 平衡：差压保护优先 / Balancing, the differential guard has priority
    eFine    := 3,    // 精抽：双泵趋近目标 / Fine pumping toward the target
    eHold    := 4,    // 保压：双腔达标保持 / Hold, both chambers at the target
    eFault   := 9     // 故障：抽速保持当前值 / Fault, the speeds keep their present values
);
END_TYPE

FUNCTION_BLOCK FB_DL_LamCtrlDualZone
VAR_INPUT
    bEnable        : BOOL := FALSE;       // 使能 / Enable
    bStartSeq      : BOOL := FALSE;       // 启动顺控，上升沿 / Start the sequence, rising edge
    fVacUpper_kPa  : REAL := 101.3;       // 上腔真空 [kPa(abs)]，域 0~101.3 / Upper chamber vacuum
    fVacLower_kPa  : REAL := 101.3;       // 下腔真空 [kPa(abs)]，域 0~101.3 / Lower chamber vacuum
    fVacTarget_kPa : REAL := 0.5;         // 目标真空 [kPa(abs)]，域 0.1~101 / Target vacuum
    fAmbient_kPa   : REAL := 101.3;       // 当地大气压 [kPa(abs)] / Local atmospheric pressure
    fDpMax_kPa     : REAL := 3.0;         // 差压上限 [kPa]，域 0.5~20 / Differential pressure limit
    fSpeedUpper    : REAL := 100.0;       // 上泵抽速给定 [%]，域 0~100 / Upper pump speed setpoint in percent
    fSpeedLower    : REAL := 100.0;       // 下泵抽速给定 [%]，域 0~100 / Lower pump speed setpoint in percent
    tSegMax        : TIME := T#60S;       // 各段超时 [ms]，域 1~600 s / Per-segment timeout
END_VAR
VAR_OUTPUT
    bVacOk         : BOOL;                // 双腔达标（双侧都不高于目标） / Both chambers at or below the target
    fDp_kPa        : REAL;                // 实时差压（上减下）[kPa] / Differential pressure, upper minus lower
    uSeg           : UINT;                // 当前段 1 粗抽 2 平衡 3 精抽 4 保压 0 待机 9 故障 [—] / Current segment
    fSpeedUpCmd    : REAL;                // 上泵指令 [%] / Upper pump command in percent
    fSpeedLowCmd   : REAL;                // 下泵指令 [%] / Lower pump command in percent
    bDpGuardActive : BOOL;                // 差压保护介入 / Differential guard active
    eErr           : UDINT;               // 错误码，段位 16#0003_xxxx / Error code in segment 16#0003_xxxx
END_VAR
VAR
    _eSeg          : E_DL_LamSeg := E_DL_LamSeg.eIdle; // 当前段 / Current segment
    _bInit         : BOOL := FALSE;       // 首扫标志，取非判定 / First-scan flag, tested negated
    _bCfgOk        : BOOL;                // 组态合法标志 / Configuration valid flag
    _bUpOk         : BOOL;                // 上腔读数有限 / Upper reading finite
    _bLowOk        : BOOL;                // 下腔读数有限 / Lower reading finite
    _fUp           : REAL;                // 上腔生效值（非有限按 0）[kPa(abs)] / Effective upper value
    _fLow          : REAL;                // 下腔生效值（非有限按 0）[kPa(abs)] / Effective lower value
    _fSpeedUp      : REAL := 100.0;       // 上泵内部指令 [%] / Internal upper command
    _fSpeedLow     : REAL := 100.0;       // 下泵内部指令 [%] / Internal lower command
    _fSegSec       : REAL;                // 段超时换算秒 [s] / Segment timeout in seconds
    _rtrigStart    : R_TRIG;              // 启动上升沿 / Rising edge of the start command
    _tonSeg        : TON;                 // 段超时计时 / Segment timeout timer
END_VAR
VAR CONSTANT
    DL_LAM_READY   : UDINT := 16#0003_03BB;  // 就绪码 / Ready code
    DL_LAM_DP_BAD  : UDINT := 16#0003_03BC;  // 故障级差压上限非法码 / Fault code for an invalid limit
    DL_LAM_TGT_BAD : UDINT := 16#0003_03BD;  // 故障级目标不可达码 / Fault code for an unreachable target
    DL_LAM_SEG_TO  : UDINT := 16#0003_03BE;  // 故障级段超时码 / Fault code for a segment timeout
    DL_LAM_SIDE_BAD : UDINT := 16#0003_03BF; // 故障级单侧非有限码 / Fault code for a non-finite side
    DL_LAM_DP_LO   : REAL := 0.5;            // 差压上限下限 [kPa] / Differential limit lower bound
    DL_LAM_DP_HI   : REAL := 20.0;           // 差压上限上限 [kPa] / Differential limit upper bound
    DL_LAM_TGT_LO  : REAL := 0.1;            // 目标真空下限 [kPa(abs)] / Target lower bound
    DL_LAM_SPD_MIN : REAL := 20.0;           // 差压保护降速后的保底抽速 [%] / Minimum speed kept by the guard
    DL_LAM_BAL_K   : REAL := 2.0;            // 平衡相触发倍率（压力 ≤ 倍率×目标即转平衡） / Balancing trigger factor
END_VAR

// 段 1｜输出与单拍标志预置
bVacOk := FALSE;                                    // 达标标志预清 / Target-reached flag pre-cleared
bDpGuardActive := FALSE;                            // 差压保护标志预清 / Guard flag pre-cleared
eErr := 0;                                          // 错误码预清 / Error code pre-cleared

// 段 2｜沿检测与段超时定时器无条件周期刷新
_rtrigStart(CLK := bStartSeq);                      // 启动沿 / Start edge
_tonSeg(IN := (_eSeg <> E_DL_LamSeg.eIdle) AND (_eSeg <> E_DL_LamSeg.eHold) AND (_eSeg <> E_DL_LamSeg.eFault), PT := tSegMax);

// 段 3｜首扫初始化（判据取非，R19）
IF NOT _bInit THEN
    _eSeg := E_DL_LamSeg.eIdle;                     // 段待机起步 / Segment starts idle
    _bInit := TRUE;                                 // 首扫只做一次 / The first scan runs once
END_IF

// 段 4｜组态闸（差压上限判零防除零；目标必须低于大气压）
_bCfgOk := NOT ((fDpMax_kPa <> fDpMax_kPa) OR ((fDpMax_kPa - fDpMax_kPa) <> (fDpMax_kPa - fDpMax_kPa)))
        AND (fDpMax_kPa >= DL_LAM_DP_LO) AND (fDpMax_kPa <= DL_LAM_DP_HI)
        AND (fVacTarget_kPa >= DL_LAM_TGT_LO)
        AND NOT ((fVacTarget_kPa <> fVacTarget_kPa) OR ((fVacTarget_kPa - fVacTarget_kPa) <> (fVacTarget_kPa - fVacTarget_kPa)))
        AND (fAmbient_kPa > 0.0);
IF _bCfgOk AND (fVacTarget_kPa >= fAmbient_kPa) THEN
    eErr := DL_LAM_TGT_BAD;                         // 故障级：目标不可达（≥ 大气压） / Fault, the target is unreachable
    _eSeg := E_DL_LamSeg.eFault;
ELSIF NOT _bCfgOk THEN
    eErr := DL_LAM_DP_BAD;                          // 故障级：差压上限非法 / Fault, the differential limit is invalid
    _eSeg := E_DL_LamSeg.eFault;
END_IF

// 段 5｜单侧读数闸（非有限侧按 0 = 最好真空；双侧齐发则停车保压）
_bUpOk := NOT ((fVacUpper_kPa <> fVacUpper_kPa) OR ((fVacUpper_kPa - fVacUpper_kPa) <> (fVacUpper_kPa - fVacUpper_kPa)));
_bLowOk := NOT ((fVacLower_kPa <> fVacLower_kPa) OR ((fVacLower_kPa - fVacLower_kPa) <> (fVacLower_kPa - fVacLower_kPa)));
IF _bUpOk THEN
    _fUp := fVacUpper_kPa;                          // 上腔有效值 [kPa(abs)] / Effective upper value
ELSE
    _fUp := 0.0;                                    // 上腔按 0（保守：视为最好真空）/ Upper side treated as zero, the conservative assumption
    eErr := DL_LAM_SIDE_BAD;                        // 故障级：上腔非有限 / Fault, the upper reading is not finite
END_IF
IF _bLowOk THEN
    _fLow := fVacLower_kPa;                         // 下腔有效值 [kPa(abs)] / Effective lower value
ELSE
    _fLow := 0.0;                                   // 下腔按 0 / Lower side treated as zero
    eErr := DL_LAM_SIDE_BAD;                        // 故障级：下腔非有限 / Fault, the lower reading is not finite
END_IF
IF (NOT _bUpOk) AND (NOT _bLowOk) THEN
    _fSpeedUp := 0.0;                               // 双侧非有限：上泵停车 [%] / Both sides invalid, the upper pump stops
    _fSpeedLow := 0.0;                              // 双侧非有限：下泵停车 [%] / Both sides invalid, the lower pump stops
    _eSeg := E_DL_LamSeg.eFault;
END_IF

// 段 6｜差压求取与保护（只降抽得快的一侧）
fDp_kPa := _fUp - _fLow;                            // 差压 = 上 − 下 [kPa] / Differential pressure
IF ABS(fDp_kPa) > fDpMax_kPa THEN
    bDpGuardActive := TRUE;                         // 差压保护介入 / The guard intervenes
    IF _fUp < _fLow THEN
        _fSpeedUp := MAX(DL_LAM_SPD_MIN, _fSpeedUp * 0.5);   // 上腔抽得快：降上泵 [%] / The upper chamber pumps faster, slow it down
    ELSE
        _fSpeedLow := MAX(DL_LAM_SPD_MIN, _fSpeedLow * 0.5); // 下腔抽得快：降下泵 [%] / The lower chamber pumps faster, slow it down
    END_IF
END_IF

// 段 7｜失能闸
IF NOT bEnable THEN
    _eSeg := E_DL_LamSeg.eIdle;                     // 段回待机 / Segment back to idle
    _fSpeedUp := 0.0;                               // 上泵指令 0 [%] / Upper command zeroed
    _fSpeedLow := 0.0;                              // 下泵指令 0 [%] / Lower command zeroed
    eErr := DL_LAM_READY;                           // 失能为正常停机 / Disable is a normal stop
END_IF

// 段 8｜双腔达标判据（双侧都不高于目标）
bVacOk := (_fUp <= fVacTarget_kPa) AND (_fLow <= fVacTarget_kPa) AND _bUpOk AND _bLowOk;

// 段 9｜四段顺控（ENUM + CASE + ELSE 兜底）
IF bEnable THEN
    CASE _eSeg OF

        E_DL_LamSeg.eIdle:                          // 待机：启动沿开粗抽
            _fSpeedUp := 0.0;
            _fSpeedLow := 0.0;
            IF _rtrigStart.Q THEN
                _fSpeedUp := LIMIT(0.0, fSpeedUpper, 100.0);   // 上泵按给定 [%] / Upper pump at the setpoint
                _fSpeedLow := LIMIT(0.0, fSpeedLower, 100.0);  // 下泵按给定 [%] / Lower pump at the setpoint
                _eSeg := E_DL_LamSeg.eRough;                   // 进入粗抽 / Enter rough pumping
            END_IF

        E_DL_LamSeg.eRough:                         // 粗抽：任一侧到 2×目标即转平衡
            IF (_fUp <= (fVacTarget_kPa * DL_LAM_BAL_K)) OR (_fLow <= (fVacTarget_kPa * DL_LAM_BAL_K)) THEN
                _eSeg := E_DL_LamSeg.eBalance;
            ELSIF _tonSeg.Q THEN
                eErr := DL_LAM_SEG_TO;              // 故障级：粗抽段超时（抽速保持） / Fault, the rough segment timed out
                _eSeg := E_DL_LamSeg.eFault;
            END_IF

        E_DL_LamSeg.eBalance:                       // 平衡：差压回到限内即转精抽
            _fSpeedUp := MAX(_fSpeedUp, DL_LAM_SPD_MIN);       // 平衡段保底抽速 [%] / Minimum speed while balancing
            _fSpeedLow := MAX(_fSpeedLow, DL_LAM_SPD_MIN);
            IF ABS(fDp_kPa) <= fDpMax_kPa THEN
                _eSeg := E_DL_LamSeg.eFine;
            ELSIF _tonSeg.Q THEN
                eErr := DL_LAM_SEG_TO;              // 故障级：平衡段超时 / Fault, the balancing segment timed out
                _eSeg := E_DL_LamSeg.eFault;
            END_IF

        E_DL_LamSeg.eFine:                          // 精抽：双腔达标即保压
            _fSpeedUp := MAX(_fSpeedUp, DL_LAM_SPD_MIN);
            _fSpeedLow := MAX(_fSpeedLow, DL_LAM_SPD_MIN);
            IF bVacOk THEN
                _eSeg := E_DL_LamSeg.eHold;
            ELSIF _tonSeg.Q THEN
                eErr := DL_LAM_SEG_TO;              // 故障级：精抽段超时 / Fault, the fine segment timed out
                _eSeg := E_DL_LamSeg.eFault;
            END_IF

        E_DL_LamSeg.eHold:                          // 保压：保持当前抽速，达标仍然成立
            IF NOT bVacOk THEN
                _eSeg := E_DL_LamSeg.eFine;         // 真空劣化：回精抽 / Vacuum degraded, back to fine pumping
            END_IF

        E_DL_LamSeg.eFault:                         // 故障：抽速保持当前值（不归零）
            eErr := DL_LAM_SEG_TO;                  // 故障级：故障段以段超时码承载 / The fault segment is carried by the timeout code
            IF _rtrigStart.Q THEN
                _fSpeedUp := LIMIT(0.0, fSpeedUpper, 100.0);   // 重启：按给定恢复 [%] / Restart restores the setpoint
                _fSpeedLow := LIMIT(0.0, fSpeedLower, 100.0);
                _eSeg := E_DL_LamSeg.eRough;
            END_IF

        ELSE
            // 非法段兜底（故障级，差压上限码承载）
            eErr := DL_LAM_DP_BAD;                  // 故障级：非法段值 / Fault, illegal segment value
            _eSeg := E_DL_LamSeg.eFault;
    END_CASE
END_IF

uSeg := 0;                                     // 段出口预置 / Segment output pre-set
CASE _eSeg OF
    E_DL_LamSeg.eIdle:    uSeg := 0;                // 待机 / Idle
    E_DL_LamSeg.eRough:   uSeg := 1;                // 粗抽 / Rough
    E_DL_LamSeg.eBalance: uSeg := 2;                // 平衡 / Balance
    E_DL_LamSeg.eFine:    uSeg := 3;                // 精抽 / Fine
    E_DL_LamSeg.eHold:    uSeg := 4;                // 保压 / Hold
    E_DL_LamSeg.eFault:   uSeg := 9;                // 故障 / Fault
    ELSE
        uSeg := 9;                                  // 非法段按故障段出口 / Illegal segments are reported as fault
END_CASE
fSpeedUpCmd := _fSpeedUp;                           // 上泵指令出口 [%] / Upper command output
fSpeedLowCmd := _fSpeedLow;                         // 下泵指令出口 [%] / Lower command output
END_FUNCTION_BLOCK

(* ---- FB_DL_LamDoorInterlock.st ---- *)
// =====================================================================
// FB_DL_LamDoorInterlock.st
// 层压机炉门-真空-温度三联锁（开门三条件 + 反向联锁 + 首因定位）
// Laminator door-vacuum-temperature interlock FB
// 码位: 16#0003_03CF ~ 16#0003_03D3 (本件独占 5 槽)
// 修改记录: R29 初版 (按 DISPATCH_R29 序 10)
// =====================================================================
FUNCTION_BLOCK FB_DL_LamDoorInterlock
VAR_INPUT
    bEnable      : BOOL  := FALSE;    // 使能 / Enable
    bReset       : BOOL  := FALSE;    // 复位 / Reset
    bDoorClosed  : BOOL  := FALSE;    // 门关到位 / Door closed
    bDoorLocked  : BOOL  := FALSE;    // 门锁定反馈 / Door locked
    bUnlockReq   : BOOL  := FALSE;    // 开门请求 / Unlock request
    bVacReleased : BOOL  := FALSE;    // 真空已破（常开触点语义外置）/ Vacuum released
    bVacReady    : BOOL  := FALSE;    // 真空泵就绪 / Vacuum pump ready
    fVac_kPa     : REAL  := 101.3;    // 腔体绝压 0~101.3 kPa / Chamber pressure [kPa]
    fTemp_C      : REAL  := 25.0;     // 腔体温度 -20~250 ℃ / Chamber temperature [degC]
    fTempSafe_C  : REAL  := 60.0;     // 允许开门温度 20~120 ℃ / Safe unlock temperature [degC]
    fHeatPct     : REAL  := 0.0;      // 加热输出 0~100 % / Heater output [%]
    tUnlockHold  : TIME  := T#5S;     // 解锁保持超时监控 T#500MS~T#60S / Unlock hold timeout [s]
END_VAR
VAR_OUTPUT
    bDoorRelease : BOOL;              // 门解锁输出 / Door release
    bHeatPermit  : BOOL;              // 允许加热 / Heat permit
    bVacPermit   : BOOL;              // 允许抽真空 / Vacuum permit
    uFirstCause  : USINT;             // 首因码 0=无 1=真空 2=温度 3=加热 4=门信号 / First cause
    bHoldTimeout : BOOL;              // 解锁保持超时 / Unlock hold timeout
    eErr         : UDINT;             // 错误码 / Error code
END_VAR
VAR
    tonHold      : TON;               // 解锁保持超时定时器（无条件周期刷新）/ Unlock hold timer
    tonExempt    : TON;               // 门信号矛盾豁免窗口定时器 / Door-signal exemption timer
    bDoorMismatch: BOOL;              // 门信号矛盾当前值 / Door mismatch current
    bMismatchLatch: BOOL := FALSE;    // 门信号矛盾故障锁存 / Door mismatch fault latch
    bVacOK       : BOOL;              // 条件 1：真空已破 / Cond 1: vacuum released
    bTempOK      : BOOL;              // 条件 2：温度安全 / Cond 2: temp safe
    bHeatOK      : BOOL;              // 条件 3：加热已撤 / Cond 3: heat off
    tHoldS       : REAL;              // 超时秒值 / Hold timeout seconds [s]
    xFirstScan   : BOOL  := TRUE;     // 首扫标记 / First-scan flag
END_VAR

// ---------------------------------------------------------------------
// 代码位表（本件独占，勿复用）:
//   16#0003_03CF 信息 联锁判定正常
//   16#0003_03D0 故障 温度/压力非有限 / tUnlockHold 非法
//   16#0003_03D1 故障 fTempSafe_C 出域（<20 或 >120）/ fVac_kPa < 0（组态错）
//   16#0003_03D2 信息 解锁保持超时（放行后门未开）→ bHoldTimeout=TRUE，不撤放行
//   16#0003_03D3 故障 bDoorClosed ≠ bDoorLocked（矛盾）→ 禁止加热/抽真空，锁存；解除=bReset 且信号一致
// ---------------------------------------------------------------------

// ---- 超时秒值 / Hold timeout seconds ----
tHoldS := TIME_TO_REAL(tUnlockHold) / 1000.0;   // 秒值 / Seconds [s]

// ---- 非有限与超时合法性闸 / Finite and timeout validity gate ----
IF (tUnlockHold = T#0MS) OR (tHoldS < 0.5) OR (tHoldS > 60.0)
   OR (fTemp_C <> fTemp_C) OR (ABS(fTemp_C) >= 1.0E12)
   OR (fVac_kPa <> fVac_kPa) OR (ABS(fVac_kPa) >= 1.0E12)
   OR (fHeatPct <> fHeatPct) OR (ABS(fHeatPct) >= 1.0E12)
   OR (fTempSafe_C <> fTempSafe_C) OR (ABS(fTempSafe_C) >= 1.0E12) THEN
    bDoorRelease := FALSE;      // 解锁输出撤销（安全侧）/ Release off (safe side)
    bHeatPermit  := FALSE;      // 加热许可撤销 / Heat permit off
    bVacPermit   := FALSE;      // 真空许可撤销 / Vac permit off
    eErr         := 16#0003_03D0;   // 故障码 / Fault code
    RETURN;                     // 本拍结束 / End of cycle
END_IF

// ---- 组态错闸 / Configuration fault gate ----
IF (fTempSafe_C < 20.0) OR (fTempSafe_C > 120.0) OR (fVac_kPa < 0.0) THEN
    bDoorRelease := FALSE;      // 解锁输出撤销 / Release off
    bHeatPermit  := FALSE;      // 加热许可撤销 / Heat permit off
    bVacPermit   := FALSE;      // 真空许可撤销 / Vac permit off
    eErr         := 16#0003_03D1;   // 故障码 / Fault code
    RETURN;                     // 本拍结束 / End of cycle
END_IF

// ---- 首扫初始化（R16 首扫纪律）/ First-scan initialization ----
IF xFirstScan THEN
    bDoorRelease := FALSE;      // 解锁初始关 / Release init off
    bHeatPermit  := FALSE;      // 加热许可初始关 / Heat permit init off
    bVacPermit   := FALSE;      // 真空许可初始关 / Vac permit init off
    xFirstScan := FALSE;        // 清标记 / Clear flag
END_IF

// ---- 使能撤销：三输出全 FALSE（安全侧）/ Disable: all outputs FALSE ----
IF NOT bEnable THEN
    bDoorRelease := FALSE;      // 解锁撤销 / Release off
    bHeatPermit  := FALSE;      // 加热撤销 / Heat off
    bVacPermit   := FALSE;      // 真空撤销 / Vac off
    bHoldTimeout := FALSE;      // 超时复位 / Timeout reset
    bMismatchLatch := FALSE;    // 锁存复位 / Latch reset
    uFirstCause  := 0;          // 首因清零 / Cause cleared
    eErr := 16#0003_03CF;       // 信息级：空闲正常 / Info: idle normal
    RETURN;                     // 本拍结束 / End of cycle
END_IF

// ---- 门信号矛盾检测（豁免窗口内不判故障）/ Door mismatch detection with exemption window ----
bDoorMismatch := (bDoorClosed <> bDoorLocked);  // 矛盾当前值 / Mismatch current
IF bDoorMismatch AND bUnlockReq AND (NOT bDoorClosed) THEN
    // 解锁瞬间锁反馈必然滞后 → tUnlockHold 窗口内豁免（防误锁）/ Exemption during unlock window
    tonExempt(IN := TRUE, PT := tUnlockHold);   // 豁免计时（无条件刷新）/ Exemption timing
    IF NOT tonExempt.Q THEN
        bDoorMismatch := FALSE;     // 窗口内豁免 / Exempted in window
    END_IF
ELSE
    tonExempt(IN := FALSE, PT := tUnlockHold);  // 窗口复位 / Window reset
END_IF

// ---- 门信号矛盾故障锁存与解除 / Door mismatch latch and release ----
IF bMismatchLatch THEN
    // 锁存中：禁止加热/抽真空，解锁也拒绝 / Latched: no heat/vac, no release
    bDoorRelease := FALSE;      // 解锁拒绝 / Release denied
    bHeatPermit  := FALSE;      // 加热禁止 / Heat denied
    bVacPermit   := FALSE;      // 真空禁止 / Vac denied
    uFirstCause  := 4;          // 首因：门信号 / Cause: door signal
    eErr         := 16#0003_03D3;   // 故障码回放 / Fault code replay
    IF bReset AND (NOT bDoorMismatch) THEN
        bMismatchLatch := FALSE;    // 解除锁存 / Release latch
    END_IF
    RETURN;                     // 本拍结束 / End of cycle
END_IF
IF bDoorMismatch THEN
    bMismatchLatch := TRUE;     // 置锁存 / Set latch
    bDoorRelease := FALSE;      // 解锁撤销 / Release off
    bHeatPermit  := FALSE;      // 加热禁止 / Heat denied
    bVacPermit   := FALSE;      // 真空禁止 / Vac denied
    uFirstCause  := 4;          // 首因 / Cause
    eErr         := 16#0003_03D3;   // 故障码 / Fault code
    RETURN;                     // 本拍结束 / End of cycle
END_IF

// ---- 开门三条件独立计布尔 / Three unlock conditions independently computed ----
bVacOK  := bVacReleased;        // 条件 1：真空已破 / Cond 1
bTempOK := (fTemp_C < fTempSafe_C);     // 条件 2：温度低于安全限 / Cond 2
bHeatOK := (fHeatPct < 0.5);    // 条件 3：无加热输出 / Cond 3

// ---- 首因定位：固定优先级（真空 → 温度 → 加热 → 门信号）/ First cause by fixed priority ----
uFirstCause := 0;               // 首因清零 / Cause cleared
IF bUnlockReq AND NOT (bVacOK AND bTempOK AND bHeatOK) THEN
    IF NOT bVacOK THEN
        uFirstCause := 1;       // 首因：真空未破 / Cause: vacuum
    ELSIF NOT bTempOK THEN
        uFirstCause := 2;       // 首因：温度过高 / Cause: temp
    ELSIF NOT bHeatOK THEN
        uFirstCause := 3;       // 首因：加热未撤 / Cause: heat
    ELSE
        uFirstCause := 4;       // 兜底：门信号异常 / Fallback: door signal
    END_IF
END_IF

// ---- 开门放行判定（三条件 AND）/ Release verdict (AND of three) ----
bDoorRelease := bUnlockReq AND bVacOK AND bTempOK AND bHeatOK;  // 放行 / Release

// ---- 解锁保持超时监控（放行后 tUnlockHold 内门仍未开）/ Unlock hold timeout monitor ----
bHoldTimeout := FALSE;          // 超时复位 / Reset
tonHold(IN := bDoorRelease AND (NOT bDoorClosed), PT := tUnlockHold);   // 定时器无条件刷新 / Unconditional refresh
IF tonHold.Q THEN
    bHoldTimeout := TRUE;       // 超时标志 / Timeout flag
    eErr := 16#0003_03D2;       // 信息级：保持超时（不撤放行）/ Info: timeout, release held
END_IF

// ---- 反向联锁：门未关严 → 禁止抽真空与加热 / Reverse interlock: door open blocks vac/heat ----
bVacPermit  := bDoorClosed AND bDoorLocked AND bVacReady;   // 抽真空许可 / Vac permit
bHeatPermit := bDoorClosed AND bDoorLocked;                 // 加热许可 / Heat permit

// ---- 正常码（未被超时信息级覆盖时）/ Normal code if not overridden ----
IF eErr <> 16#0003_03D2 THEN
    eErr := 16#0003_03CF;       // 信息级：联锁判定正常 / Info: normal
END_IF

END_FUNCTION_BLOCK

(* ---- FB_DL_LoadcellTareCtrl.st ---- *)
(*
  组件名 Component   : FB_DL_LoadcellTareCtrl
  子库 Sublibrary    : DL_Device
  版本 Version       : 1.0.0
  兼容性 Platform    : CODESYS 3.5 / TwinCAT 3 / 汇川 InoProShop / Machine Expert（仅 Standard.library）
  功能 Function      : 称重传感器去皮/标定管理：
                       1) 去皮锁存：bTareCmd 上升沿把当下毛重读数锁存为皮重，
                       净重 = 毛重 - 皮重（锁存量，不随后续漂移）；
                       2) 两点标定：bCalCmd 上升沿按两点已知质量与其原始读数解算
                       斜率/截距（读数跨度近零前置拦截，不进入除法）；
                       3) 标定超期计数：使能期扫描累计，超过 uCalIntervalScans 置
                       bCalDue（维护提示，信息级语义，不置 bError）；
                       4) 非有限读数判输入非法，净重出口冻结保持（安全侧）。
  边界 Boundary      : ① 本件只做称重管理，不写物理 IO（原始读数由上层适配层传入）；
                       ② 皮重/标定系数均为锁存回放，禁按当下输入重推断（R152）；
                       ③ 故障锁存解除唯一路径 = bReset 上升沿（输入引脚，恒可达）；
                       ④ Device 件无 NE107 出口（去皮/标定为维护工序件，非诊断件）；
                       ⑤ 无全局变量引用、无外部变量声明、无物理地址寻址。
  依赖 Depends       : Standard.library（R_TRIG）
  溯源 Origin        : 道莅自研 clean-room（参考 t2-6-rockwell-aoi 设备级粒度分类与
                       参数域，零代码行复制）
  码位 Code          : 16#03_2_E（Device 05xx 副带 052E）
  码表 Error codes（Device 故障窗口 052E，本件无信息码，单故障总码 + 成因枚举归因）:
    16#0003_052E 故障级：称重管理故障总码（标定读数跨度近零 / 皮重超量程 /
                 组态非法 / 输入非有限），锁存至 bReset 上升沿，归因见 eCause
  修订历史 Revision  :
    2026-11-19  v1.0.0  R44 首版（批次 2 · 序号 10）
*)

TYPE E_DL_LtcState :
(
    eIdle  := 0,    // 空闲：未使能 / Idle, not enabled
    eRun   := 10,   // 运行：去皮/标定/净重合成 / Running, tare, calibrate and net
    eFault := 90    // 故障：总码锁存 / Fault, latched
);
END_TYPE

TYPE E_DL_LtcCause :
(
    eNone      := 0,  // 无故障成因 / No cause
    eCalSpan   := 1,  // 标定读数跨度近零 / Calibration span near zero
    eTareRange := 2,  // 皮重超量程（皮重 >= 满量程） / Tare beyond capacity
    eCfgIllegal:= 3,  // 组态非法 / Illegal configuration
    eNonFinite := 4   // 输入非有限 / Non-finite input
);
END_TYPE

FUNCTION_BLOCK FB_DL_LoadcellTareCtrl
VAR_INPUT
    bEnable    : BOOL;                     // 使能（电平）[-] / Enable
    bReset     : BOOL;                     // 上升沿清故障锁存 [-] / Reset edge
    bTareCmd   : BOOL;                     // 去皮指令（上升沿承载）[-] / Tare command edge
    bCalCmd    : BOOL;                     // 标定指令（上升沿承载）[-] / Calibrate command edge
    fGrossG    : REAL;                     // 毛重读数 [克] / Gross reading
    fCalMassLoG: REAL;                     // 标定点 1 已知质量 [克] / Calibration mass 1
    fCalMassHiG: REAL;                     // 标定点 2 已知质量 [克] / Calibration mass 2
    fRawLo     : REAL;                     // 标定点 1 原始读数 [克] / Calibration raw 1
    fRawHi     : REAL;                     // 标定点 2 原始读数 [克] / Calibration raw 2
    fCapacityG : REAL := 10000.0;          // 传感器满量程 [克] / Sensor capacity
    uCalIntervalScans: UDINT := 8640000;  // 标定超期计数限 [拍] / Calibration due interval
END_VAR
VAR_OUTPUT
    fNetG      : REAL;                     // 净重输出 [克] / Net weight output
    fTareG     : REAL;                     // 锁存皮重 [克] / Latched tare weight
    fSlope     : REAL;                     // 标定斜率 [克/克读数] / Calibration slope
    fOffset    : REAL;                     // 标定截距 [克] / Calibration offset
    bTared     : BOOL;                     // 已去皮标志 [-] / Tared flag
    bCalOk     : BOOL;                     // 标定有效标志 [-] / Calibration valid flag
    bCalDue    : BOOL;                     // 标定超期标志 [-] / Calibration due flag
    uScansSinceCal: UDINT;                 // 距上次标定扫描累计 [拍] / Scans since calibration
    eState     : E_DL_LtcState;            // 状态出口，段尾单点映射 / State outlet
    eCause     : E_DL_LtcCause;            // 故障成因出口（R190） / Fault cause outlet
    bError     : BOOL;                     // 故障锁存标志 [-] / Fault latch flag
    uErrId     : UDINT;                    // 事件码，0 = 无事件 / Event code
END_VAR
VAR
    rtReset: R_TRIG;                       // 复位沿实例，段 0 无条件刷新 / Reset edge
    rtTare : R_TRIG;                       // 去皮沿实例，段 0 无条件刷新 / Tare edge
    rtCal  : R_TRIG;                       // 标定沿实例，段 0 无条件刷新 / Calibrate edge
    _eState: E_DL_LtcState := E_DL_LtcState.eIdle;     // 内部相位（CASE 唯一写入目标）/ Internal phase
    _eCause: E_DL_LtcCause := E_DL_LtcCause.eNone;     // 故障成因锁存（锁存量）/ Latched cause
    _bFault: BOOL;                         // 故障锁存位（锁存量） / Latched fault bit
    _uFault: UDINT;                        // 故障码锁存（锁存量） / Latched fault code
    _bCfgBad: BOOL;                        // 组态非法当拍量 [-] / Config illegal flag
    _bNonFin: BOOL;                        // 输入非有限当拍量 [-] / Non-finite input flag
    _bNetFin: BOOL;                        // 净重合成非有限当拍量 [-] / Net synthesis non-finite flag
    _fNetNew: REAL;                        // 净重合成暂存 [克]（过闸后才提交出口）/ Net synthesis temp
END_VAR
VAR CONSTANT
    DL_SPAN_EPS : REAL := 1.0E-6;          // 标定跨度近零判据 [克] / Span near-zero tolerance
    DL_ABS_MAX  : REAL := 1.0E30;          // 有限值判定上界 [克] / Finite bound
    DL_ZERO     : REAL := 0.0;             // 零常量 [克] / Zero constant
END_VAR

(* —— 段 0｜沿实例每拍无条件刷新（禁置于 IF/CASE 内） —— *)
rtReset(CLK := bReset);
rtTare (CLK := bTareCmd);
rtCal  (CLK := bCalCmd);

(* —— 段 1｜瞬时量预清零（锁存量 _bFault/_uFault/fTareG/fSlope/fOffset 不入清单） —— *)
uErrId   := 16#0000_0000;
_bCfgBad := FALSE;
_bNonFin := FALSE;
_bNetFin := FALSE;

(* —— 段 2｜复位沿：故障一次性清干净，相位回空闲 —— *)
IF rtReset.Q THEN
    _bFault := FALSE;
    _uFault := 16#0000_0000;
    _eCause := E_DL_LtcCause.eNone;
    _eState := E_DL_LtcState.eIdle;
END_IF

(* —— 段 3｜组态闸与非有限判据 —— *)
IF (fCapacityG <= DL_ZERO) OR (uCalIntervalScans = UDINT#0) THEN
    _bCfgBad := TRUE;
END_IF
IF (fGrossG <> fGrossG) OR ((fGrossG - fGrossG) <> DL_ZERO) THEN
    _bNonFin := TRUE;
END_IF

(* —— 段 4｜标定超期计数：使能期累计，超限置到期（信息级语义，不置 bError） —— *)
IF bEnable AND (NOT _bFault) THEN
    uScansSinceCal := uScansSinceCal + UDINT#1;
    IF uScansSinceCal >= uCalIntervalScans THEN
        bCalDue := TRUE;
    END_IF
END_IF

(* —— 段 5｜主状态机：三态全覆盖 + ELSE 兜底 —— *)
CASE _eState OF

E_DL_LtcState.eIdle:
    IF bEnable AND (NOT _bCfgBad) THEN
        _eState := E_DL_LtcState.eRun;
    ELSIF bEnable AND _bCfgBad THEN
        _bFault := TRUE;                 // 故障级配对置位（R45）
        _uFault := 16#0003_052E;
        _eCause := E_DL_LtcCause.eCfgIllegal;
        bError  := TRUE;
        _eState := E_DL_LtcState.eFault;
    END_IF

E_DL_LtcState.eRun:
    IF NOT bEnable THEN
        _eState := E_DL_LtcState.eIdle;  // 使能撤销回空闲，皮重与标定系数保持
    ELSE
        IF _bNonFin THEN
            _bFault := TRUE;             // 读数非有限：锁存，净重出口冻结保持
            _uFault := 16#0003_052E;
            _eCause := E_DL_LtcCause.eNonFinite;
            bError  := TRUE;
            _eState := E_DL_LtcState.eFault;
        ELSE
            (* 净重合成：已标定走斜率/截距链，未标定直通毛皮差；暂存过闸后才提交 *)
            IF bCalOk THEN
                _fNetNew := fSlope * fGrossG + fOffset - fTareG;
            ELSE
                _fNetNew := fGrossG - fTareG;
            END_IF
            _bNetFin := (_fNetNew <> _fNetNew) OR ((_fNetNew - _fNetNew) <> DL_ZERO)
                        OR (ABS(_fNetNew) > DL_ABS_MAX);
            IF _bNetFin THEN
                _bFault := TRUE;         // 合成结果越域/非有限：锁存，出口保持上拍值
                _uFault := 16#0003_052E;
                _eCause := E_DL_LtcCause.eNonFinite;
                bError  := TRUE;
                _eState := E_DL_LtcState.eFault;
            ELSE
                fNetG := _fNetNew;       // 过闸提交（出口单点写）
            END_IF
            (* 去皮沿：锁存当下净重前毛重为皮重，皮重超量程判非法 *)
            IF rtTare.Q AND (NOT _bFault) THEN
                IF fGrossG >= fCapacityG THEN
                    _bFault := TRUE;
                    _uFault := 16#0003_052E;
                    _eCause := E_DL_LtcCause.eTareRange;
                    bError  := TRUE;
                    _eState := E_DL_LtcState.eFault;
                ELSE
                    fTareG := fGrossG;
                    bTared := TRUE;
                END_IF
            END_IF
            (* 标定沿：两点跨度近零拦截后解算斜率/截距，标定计数清零 *)
            IF rtCal.Q AND (NOT _bFault) THEN
                IF ABS(fRawHi - fRawLo) <= DL_SPAN_EPS THEN
                    _bFault := TRUE;     // 跨度近零：斜率无意义
                    _uFault := 16#0003_052E;
                    _eCause := E_DL_LtcCause.eCalSpan;
                    bError  := TRUE;
                    _eState := E_DL_LtcState.eFault;
                ELSE
                    fSlope := (fCalMassHiG - fCalMassLoG) / (fRawHi - fRawLo);
                    fOffset := fCalMassLoG - fSlope * fRawLo;
                    bCalOk := TRUE;
                    uScansSinceCal := UDINT#0;
                    bCalDue := FALSE;
                END_IF
            END_IF
        END_IF
    END_IF

E_DL_LtcState.eFault:
    bError := TRUE;                      // 故障相驻留：净重冻结保持，只认复位沿（段 2 迁出）
    ;                                    // （冻结语义：fNetG 保持故障前值，不静默归零）

ELSE
    _bFault := TRUE;                     // 兜底：非法相位锁存
    _uFault := 16#0003_052E;
    _eCause := E_DL_LtcCause.eCfgIllegal;
    bError  := TRUE;
    _eState := E_DL_LtcState.eFault;
END_CASE

(* —— 段 6｜状态出口单点映射（名实同源） —— *)
eState := _eState;
END_FUNCTION_BLOCK

(* ---- FB_DL_MeterPulseLossDetect.st ---- *)
(*
  Name        : FB_DL_MeterPulseLossDetect
  Category    : DL_Device
  Version     : 1.0.0
  Purpose     : 脉冲式流量计丢脉冲检测：按指令流量与 K 系数推算采样窗内应有脉冲数，与实际累计脉冲增量比对，超容差即判丢脉冲；/ Detect pulse loss on a pulse-output flow meter by comparing expected pulses (command flow x K-factor) against the actual count increment within a sampling window
  溯源        : 借 t1-3-oscat-network·计量 的分类/参数域组织，clean-room 实现
  Boundary    : ① 组态闸：K 系数/采样周期/流量下限/容差任一越域 → 锁存故障；
                ② 流量闸：指令流量 <= 最小有效流量时不判（低流量下脉冲稀疏，比对无意义）；
                ③ 推算除子闸：应有脉冲数 <= eps → 不判（避免小分母放大误差）；
                ④ 累计脉冲负增量（清零/溢出回卷）按 0 处理并计入 bCountReset，不判丢脉冲；
                ⑤ 全部比值判据用容差比较，禁 `=`/`<>`。
*)
TYPE E_DL_MplState :
(
    eIdle  := 0,                             (* 未使能 / Disabled *)
    eMon   := 10,                            (* 比对运行 / Comparing *)
    eFault := 90                             (* 故障锁存相 / Fault latched *)
);
END_TYPE

TYPE E_DL_MplCause :
(
    eNone       := 0,                        (* 无故障成因 / No cause *)
    eCfgIllegal := 1,                        (* 组态非法：K 系数/周期/流量闸越域 / Illegal config *)
    ePhaseBad   := 2                         (* 非法相位兜底 / Illegal phase fallback *)
);
END_TYPE

FUNCTION_BLOCK FB_DL_MeterPulseLossDetect
VAR_INPUT
    diPulseCount : DINT := 0;                (* 流量计累计脉冲数（表侧原始累计）[脉冲] / Meter cumulative pulse count *)
    fFlowCmd     : REAL := 0.0;              (* 指令/参考流量（工艺给定），域 >= 0 [L/min] / Command (reference) flow, >= 0 *)
    fKFactor     : REAL := 100.0;            (* 仪表 K 系数（脉冲/升），域 > 0 [脉冲/L] / Meter K factor, > 0 *)
    tSample      : TIME := T#1S;             (* 采样窗长，域 > T#0S [ms] / Sampling window, > 0 *)
    fFlowMin     : REAL := 0.5;              (* 最小有效流量（判据闸），域 > 0 [L/min] / Minimum valid flow, > 0 *)
    fLossTolPct  : REAL := 10.0;             (* 丢脉冲容差，域 0 < x < 100 [%] / Loss tolerance, 0..100 *)
    bEnable      : BOOL := TRUE;             (* 检测使能 [-] / Enable *)
    bReset       : BOOL := FALSE;            (* 复位命令，上升沿清比对结果与故障 [-] / Reset command *)
END_VAR
VAR_OUTPUT
    diPulseDelta : DINT;                     (* 本窗实际脉冲增量 [脉冲] / Actual pulse increment this window *)
    fPulseExpect : REAL;                     (* 本窗应有脉冲数（推算值）[脉冲] / Expected pulses this window *)
    fLossPct     : REAL;                     (* 丢脉冲百分比（0 = 不丢，> 0 为丢失比例）[%] / Pulse loss percentage *)
    bPulseLoss   : BOOL;                     (* 丢脉冲判据（超容差）[-] / Pulse loss verdict *)
    bFlowGate    : BOOL;                     (* 流量闸开放（本窗参与判据）[-] / Flow gate open this window *)
    bCountReset  : BOOL;                     (* 累计计数回卷/清零检测位 [-] / Count reset or wrap detected *)
    eState       : E_DL_MplState;            (* 状态出口 / State outlet *)
    eCause       : E_DL_MplCause;            (* 故障成因出口（R190 归因唯一） / Fault cause outlet *)
    bError       : BOOL;                     (* 故障锁存标志 [-] / Fault latch flag *)
END_VAR
VAR
    _eState  : E_DL_MplState := E_DL_MplState.eIdle;     (* 内部相位（CASE 唯一写入目标） / Internal phase *)
    _eCause  : E_DL_MplCause := E_DL_MplCause.eNone;     (* 故障成因锁存量 / Latched cause *)
    rtReset  : R_TRIG;                       (* 复位沿实例，段 0 无条件调用 / Reset edge instance *)
    tonWin   : TON;                          (* 采样窗自复位计时器（R188） / Self-resetting window timer *)
    _bFault  : BOOL;                         (* 故障锁存位 / Latched fault bit *)
    _bCfgBad : BOOL;                         (* 组态非法当拍量 / Illegal config this scan *)
    _bFinite : BOOL;                         (* 输入有限性当拍量 / Input finiteness *)
    _diPrev  : DINT;                         (* 上窗脉冲数快照 [脉冲] / Previous window pulse snapshot *)
    _diDelta : DINT;                         (* 本窗增量（负值按 0）[脉冲] / Delta, negative treated as zero *)
    _fDtSec  : REAL;                         (* 窗长秒值 [s] / Window length in seconds *)
    _fExpect : REAL;                         (* 应有脉冲数推算中间量 [脉冲] / Expected pulses intermediate *)
    _fLoss   : REAL;                         (* 丢脉冲百分比中间量 [%] / Loss intermediate *)
END_VAR
VAR CONSTANT
    DL_MPL_EPS     : REAL := 1.0E-6;         (* 判零容差 [-] / Epsilon *)
    DL_MPL_SECMIN  : REAL := 60.0;           (* 每分秒数（L/min → L/s 换算常量）[s] / Seconds per minute *)
    DL_MPL_PCTMAX  : REAL := 100.0;          (* 百分比满量程 [%] / Percentage full scale *)
END_VAR

(* —— 段 0：当拍判据派生 + 实例无条件刷新（R228A） —— *)
_fDtSec := TIME_TO_LREAL(tSample) / 1000.0;                                    (* 窗长秒化（除子常量 1000） / Window to seconds *)
_bCfgBad := NOT (tSample > T#0S)                                               (* 窗长正域闸 / Window gate *)
            OR (fKFactor <= DL_MPL_EPS)                                        (* K 系数正域闸（乘性因子，零则无脉冲语义） / K factor gate *)
            OR (fFlowMin <= DL_MPL_EPS)                                        (* 流量闸正域 / Flow gate positive *)
            OR (fLossTolPct <= 0.0) OR (fLossTolPct >= DL_MPL_PCTMAX);         (* 容差域闸 (0,100) / Tolerance gate *)
rtReset(CLK := bReset);                                                        (* 复位沿每拍必调 / Reset edge every scan *)
tonWin(IN := NOT tonWin.Q, PT := tSample);                                     (* 采样窗自复位（R188） / Self-resetting window *)
_bFinite := (fFlowCmd = fFlowCmd) AND ((fFlowCmd - fFlowCmd) = (fFlowCmd - fFlowCmd));   (* NaN/Inf 联合闸 / NaN and Inf gate *)

(* —— 段 1：单拍量预清零（R107） —— *)
bPulseLoss := FALSE;                                                           (* 丢脉冲判据预清 / Verdict preset *)
bFlowGate := FALSE;                                                            (* 流量闸预清 / Gate preset *)
bCountReset := FALSE;                                                          (* 计数回卷位预清 / Reset flag preset *)

(* —— 段 2：复位沿处理（作用域：清故障 + 清比对 + 清快照 + 迁 eIdle，R283 逐项声明） —— *)
IF rtReset.Q THEN
    _bFault := FALSE;                                                          (* 清故障锁存 / Clear fault *)
    _eCause := E_DL_MplCause.eNone;                                            (* 清成因 / Clear cause *)
    _diPrev := diPulseCount;                                                   (* 快照对齐当前值（复位后不产生虚假增量） / Align snapshot *)
    diPulseDelta := 0;                                                         (* 清增量出口 / Clear delta *)
    fPulseExpect := 0.0;                                                       (* 清推算出口 / Clear expected *)
    fLossPct := 0.0;                                                           (* 清丢包出口 / Clear loss *)
    _eState := E_DL_MplState.eIdle;                                            (* 迁未使能相 / Back to idle *)
END_IF

(* —— 段 3：组态故障锁存（锁存至复位沿，R189） —— *)
IF _bCfgBad AND NOT _bFault THEN
    _bFault := TRUE;                                                           (* 锁存故障位 / Latch fault *)
    _eCause := E_DL_MplCause.eCfgIllegal;                                      (* 成因：组态非法 / Cause: illegal config *)
    _eState := E_DL_MplState.eFault;                                           (* 同步迁故障相 / Migrate to fault *)
END_IF

(* —— 段 4：CASE 主状态机（ELSE 兜底迁 eFault，红线 6） —— *)
CASE _eState OF
    E_DL_MplState.eIdle:                                                       (* 未使能：快照持续跟随，不判 / Disabled *)
        _diPrev := diPulseCount;                                               (* 失能期间跟随（重使能无虚假增量） / Track while disabled *)
        IF bEnable AND NOT _bFault THEN
            _eState := E_DL_MplState.eMon;                                     (* 使能进入比对 / Enter comparing *)
        END_IF
    E_DL_MplState.eMon:                                                        (* 比对相：窗到点结算一次 / Comparing *)
        IF NOT bEnable THEN
            _eState := E_DL_MplState.eIdle;                                    (* 失能回未使能 / Back to idle *)
        ELSIF tonWin.Q THEN                                                    (* 窗到点：单点结算 / Window elapsed: settle once *)
            _diDelta := diPulseCount - _diPrev;                                (* 增量 = 当前 - 上窗快照 / Delta *)
            IF _diDelta < 0 THEN
                _diDelta := 0;                                                 (* 负增量（清零/回卷）：按 0 处理 / Negative: zero *)
                bCountReset := TRUE;                                           (* 标记计数回卷，不判丢脉冲（边界④） / Mark wrap, skip verdict *)
            END_IF
            diPulseDelta := _diDelta;                                          (* 增量出口 / Delta outlet *)
            _diPrev := diPulseCount;                                           (* 快照推进（单点写入，无双向双计） / Advance snapshot *)
            IF _bFinite AND (fFlowCmd > fFlowMin) THEN                         (* 流量闸：低流量不判 / Flow gate *)
                bFlowGate := TRUE;                                             (* 闸开放 / Gate open *)
                _fExpect := fFlowCmd / DL_MPL_SECMIN * _fDtSec * fKFactor;     (* 应有脉冲 = (L/min→L/s)·s·K（除子为常量）[脉冲] / Expected pulses *)
                fPulseExpect := _fExpect;                                      (* 推算出口 / Expected outlet *)
                IF _fExpect > DL_MPL_EPS THEN                                  (* 除子闸（边界③） / Divisor gate *)
                    _fLoss := (1.0 - DINT_TO_REAL(_diDelta) / _fExpect) * DL_MPL_PCTMAX;   (* 丢脉冲百分比（除子已过闸）[%] / Loss percentage *)
                    IF _fLoss < 0.0 THEN
                        _fLoss := 0.0;                                         (* 多计数（负丢包）按 0 饱和 / Clamp to zero *)
                    ELSIF _fLoss > DL_MPL_PCTMAX THEN
                        _fLoss := DL_MPL_PCTMAX;                               (* 上限饱和 100% / Upper saturation *)
                    END_IF
                    fLossPct := _fLoss;                                        (* 丢包出口 / Loss outlet *)
                    IF _fLoss > fLossTolPct THEN
                        bPulseLoss := TRUE;                                    (* 超容差：判丢脉冲 / Exceeds tolerance: loss *)
                    END_IF
                ELSE
                    fLossPct := 0.0;                                           (* 推算量过小：不判，出口清 0 / Too small: no verdict *)
                END_IF
            ELSE
                bFlowGate := FALSE;                                            (* 闸关闭：本窗不判 / Gate closed *)
                fPulseExpect := 0.0;                                           (* 推算出口清 0（无判据语义） / Expected cleared *)
                fLossPct := 0.0;                                               (* 丢包出口清 0 / Loss cleared *)
            END_IF
        END_IF
    E_DL_MplState.eFault:                                                      (* 故障相：冻结保持末值，仅复位沿出 / Fault *)
        ;                                                                      (* 锁存回放（R28） / Replay from latch *)
    ELSE                                                                       (* 非法相位兜底迁安全态 / Illegal phase fallback *)
        _eState := E_DL_MplState.eFault;                                       (* 迁故障相 / To fault *)
        _bFault := TRUE;                                                       (* 同步锁存 / Latch *)
        _eCause := E_DL_MplCause.ePhaseBad;                                    (* 成因：非法相位 / Cause: illegal phase *)
END_CASE

(* —— 段 5：出口映射（bError/eState 同源，R191） —— *)
bError := _bFault;                                                             (* 故障标志镜像 / Fault flag mirror *)
eState := _eState;                                                             (* 状态出口 / State outlet *)
eCause := _eCause;                                                             (* 成因出口 / Cause outlet *)
END_FUNCTION_BLOCK
